FUNCTION_BLOCK FTS_NCGenerator
VAR_IN_OUT
	stAxis: ST_Axis;
END_VAR
VAR_INPUT
	///滤波窗口大小
	nWindowSize: UINT;
	fCycleTime: LREAL;
END_VAR
VAR
	///_bCalStart             :BOOL:=FALSE;
	_bEnable: BOOL;
	///_bAutoPlan             :BOOL:=FALSE;
	_bCalculateDone: BOOL;
	_bSynMode: BOOL := FALSE;
	_bFisrtUpdate: BOOL := FALSE;
	_bEndOfProfile: BOOL := FALSE;
	_bEstopping: BOOL := FALSE;
	///03.31     
	_bIsGroupMember: BOOL := FALSE;
	_bAddNodeOk: BOOL := FALSE;
	_bDeleteNodeOk: BOOL := FALSE;
	_bInsertOk: BOOL := FALSE;
	_bPreEstop  :BOOL:=FALSE;
	_bPreDyEstop  :BOOL:=FALSE;
	_nIndex: INT;
	_nNodeIndex: UINT;
	_nLastIndex: INT;
	_nPointIndex: UINT;
	_nForwardIndex: INT;
	_nPreIndex: INT;
	_nState: INT;
	_nPathSegment: INT;
	_nSysType: UINT;
	_nCamBufferNum: UINT := 0;
	_nCuRoadID: UINT;
	_nLastRoadID: UINT;
	_nMoverCounter: UINT;
	_nLastMoverCounter: UINT;
	_fRealDis: LREAL;
	_fPos: LREAL;
	_fSynPos: LREAL;
	_fSynVelo: LREAL;
	_lastVelo: LREAL;
	_fVeloStart: LREAL;
	_fVeloEnd: LREAL;
	_fTargetVelo: LREAL;
	_fStartPos: LREAL;
	_fEndPos: LREAL;
	_fVeloStart_2: LREAL;
	_fVeloEnd_2: LREAL;
	_fTargetVelo_2: LREAL;
	_fDistance_2: LREAL;
	_fAcc: LREAL;
	_fDec: LREAL;
	_fJerk: LREAL;
	_fAcc_2: LREAL;
	_fDec_2: LREAL;
	_fDistance: LREAL;
	///_fDistance_2             :LREAL;
	_fSetVelo: LREAL;
	///夹具长度*0.5
	_fGap: LREAL;
	_fGapSet: LREAL;
	_fTime: LREAL;
	_fDisSet: LREAL;
	_fForwardTime: LREAL;
	_fDealtDis: LREAL;
	_fDealt_S: LREAL;
	_fPre_S: LREAL;
	_fPreDealt_S: LREAL;
	_fDealt_S1: LREAL;
	_fPreCuVel: LREAL;
	_fCuVel: LREAL;
	_fPreTaVel: LREAL;
	_fPreAcc: LREAL;
	_fNewAcc: LREAL;
	_fDecTime: LREAL;
	_fDecTime_1: LREAL;
	_fPreCurTime: LREAL;
	_fPreSeg1TotalTime: LREAL;
	_fDisDiff: LREAL;
	_fDealDecTime: LREAL;
	_fMinDis: LREAL;
	_fNewAccDis: LREAL;
	_fReminDis: LREAL;
	_fAccMisDis: LREAL;
	_fAccMisDis_1: LREAL;
	_fNewVelo: LREAL;
	_fStartLinearPos: LREAL;
	_fLinearDealt: LREAL;
	_fMasterPos: LREAL;
	_fMasterStartPos: LREAL;
	_fMasterEndPos: LREAL;
	_fSlaveStartPos: LREAL;
	_fDePos: LREAL;
	_fDeCuVelo: LREAL;
	_fVeloRatio: LREAL;
	_fPos_X: LREAL;
	_fDealt_X: LREAL;
	_fLastPos: LREAL;
	_fMasterGap: LREAL;
	_fRoad1_Lenth: LREAL;
	_fRoad2_Lenth: LREAL;
	_fCuRoadLenth: LREAL;
	_fPosTemp: LREAL;
	_fLastPosDeat: LREAL;
	_fLastPosNC: LREAL;
	_fPosIn: LREAL;
	_fStopPos: LREAL;
	_fEStopPos: LREAL;
	_fPreStopPos: LREAL;
	_fUpNewPos: LREAL;
	_fUpNewPosTemp: LREAL;
	/// 成组组内gap 03.31
	_fGroupInGap: LREAL;
	///06.30
	_fSetDealtGap: LREAL;
	_fPyRealdis  :LREAL; //02.28
	_fLastRoadPos :LREAL;
	_fBreakDis    :LREAL;   
	_fSetSafeDis  :LREAL;
	_fLastPtyPos  :LREAL;
	_fPtyVelo    :LREAL;
	
	_fPreDealtP  :LREAL;
	
	///_fEndPos               :LREAL;  //03.26
	_sMessage3: STRING;
	_sMessage: STRING(1024);
	_sMessage2: STRING(1024);
	
	_pPremover: POINTER TO ST_Axis;
	_pNextRoadPremover: POINTER TO ST_Axis;
	///_fStopTime             :LREAL;
	_ePlanningMode: E_PlanningMode;
	_stAxis_Point: ST_Point;
	_stLastAxis_Point: ST_Point;
	_stForwardAxis_Point: ST_Point;
	_stPreAxis_Point: ST_Point;
	_stAxisNo: ST_Axis;
	_eDirection: E_Direction;
	///04.08
	_eSetDirection: E_Direction;
	_stTimeInfo: ST_TimeRef;
	_stTimeInfo_2: ST_TimeRef;
	_stPathRef: ST_PathRef;
	_stNoPathRef: ST_PathRef;
	_stPolynom5Factor: ST_Polynom5Factor;
	_stSShapedParam: ST_SParam;
	_stCamParam: ST_CamParam;
	_aLinearPosition: ARRAY[1..100] OF LREAL;
	_aCamBuffer: ARRAY[0..9] OF ST_CamXYVA;
	_fbTrig: R_TRIG;
	_fbSlaveTrig: R_TRIG;
	_fbPathTrig: R_TRIG;
	_fbDecPathTrig: R_TRIG;
	_fbCamPointUpdateTrig: R_TRIG;
	_fbCamBufUpdateTrig: R_TRIG;
	_fbClearFtrig: F_TRIG;
	_fbDecNextPathTrig: R_TRIG;
	_fbAxis: FB_TrajectoryPlanning;
	_fbPreAxis: FB_TrajectoryPlanning;
	_fbTon: TON;
	_fbFilterV2: FB_FilterWindowV2;
	_fbStopTrig: R_TRIG;
	_fbStopTon: TON;
	_fbAxisGroupList: FTS_AxisGroupList;
	_fbTrigRoadUpdate: R_TRIG;
	_fbTrigRoadDeleUpdate: R_TRIG;
	_fbTonCuPos:ton ; //02.28
END_VAR
VAR CONSTANT
	//cDebug: BOOL := TRUE;
	cStateIdle: INT := 0;
	cStateReady: INT := 1;
	cStatePathGenerator: INT := 2;
	cDealtGap: REAL := 10000;
	//cNcCycle: REAL := 0.001;
	cPointBuffer: UINT := 10;
END_VAR


// control logic 
IF stAxis.stAxisStatus.bPositiveDirection THEN 
	_eDirection:=E_Direction.DIRECTION_POSITIVE;
	
ELSIF stAxis.stAxisStatus.bNegativeDirection  THEN
	_eDirection:=E_Direction.DIRECTION_NEGATIVE;
	
ELSE
	_eDirection:=E_Direction.DIRECTION_POSITIVE;
END_IF

//根据不同road 前置和后置配置  04/02
IF (stAxis.stPLCTONC.nRoadID_2<>0)AND (stAxis.stPLCTONC.nRoadID_1<>0)AND(stAxis.stNcTOPLC.nCuRoadID=stAxis.stPLCTONC.nRoadID_2)THEN   //04.02
	
		IF NOT stAxis.stPLCTONC.bRoadDirection  THEN
			IF (stAxis.stAxisStatus.pPremover=0)THEN 
				_pPremover:=ADR(_stAxisNo);
			ELSE
				_pPremover:=stAxis.stAxisStatus.pPremover;
			END_IF
		ELSE
			IF (stAxis.stAxisStatus.pAftermover=0)THEN 
				_pPremover:=ADR(_stAxisNo);
			ELSE
				_pPremover:=stAxis.stAxisStatus.pAftermover;
			END_IF
		END_IF	
ELSE
	IF (_eDirection=E_Direction.DIRECTION_POSITIVE)THEN 
		IF (stAxis.stAxisStatus.pPremover=0)THEN 
			_pPremover:=ADR(_stAxisNo);
		ELSE
			_pPremover:=stAxis.stAxisStatus.pPremover;
		END_IF
	ELSE
		IF (stAxis.stAxisStatus.pAftermover=0)THEN 
			_pPremover:=ADR(_stAxisNo);
		ELSE
			_pPremover:=stAxis.stAxisStatus.pAftermover;
		END_IF
	
	END_IF
END_IF

IF (stAxis.stAxisStatus.pNextRoadPremover=0)THEN
	_pNextRoadPremover :=ADR(_stAxisNo);
ELSE
	_pNextRoadPremover :=stAxis.stAxisStatus.pNextRoadPremover;
END_IF

// 是否成组判断，并根据条件计算组内gap距离  03.31
IF (_pPremover^.stNcTOPLC.nAxisId<>0) THEN 
	IF (_pPremover^.stAxisStatus.stGroupRef.eGroupType<>E_GroupType.GROUPTYPE_NONE)
           AND (stAxis.stAxisStatus.stGroupRef.eGroupType<>E_GroupType.GROUPTYPE_NONE)THEN 
		IF (_pPremover^.stAxisStatus.stGroupRef.nGroupId=stAxis.stAxisStatus.stGroupRef.nGroupId)THEN 
			//_fGroupInGap:=stAxis.stAxisStatus.stPathRef.fGroupInGap;
			_fGroupInGap:=stAxis.stPLCTONC.fGroupInGap;
			_bIsGroupMember:=TRUE;
		END_IF
	ELSE
		_bIsGroupMember:=FALSE;
	END_IF
ELSE
	IF (_pNextRoadPremover^.stNcTOPLC.nAxisId<>0) THEN 
		IF (_pNextRoadPremover^.stAxisStatus.stGroupRef.eGroupType<>E_GroupType.GROUPTYPE_NONE)
			   AND (stAxis.stAxisStatus.stGroupRef.eGroupType<>E_GroupType.GROUPTYPE_NONE)THEN 
			IF (_pNextRoadPremover^.stAxisStatus.stGroupRef.nGroupId=stAxis.stAxisStatus.stGroupRef.nGroupId)THEN 
				//_fGroupInGap:=stAxis.stAxisStatus.stPathRef.fGroupInGap;
				_fGroupInGap:=stAxis.stPLCTONC.fGroupInGap;
				_bIsGroupMember:=TRUE;
			END_IF
		ELSE
			_bIsGroupMember:=FALSE;
		END_IF
	ELSE 
	   _bIsGroupMember:=FALSE;
	END_IF
END_IF



// 前后动子实时位置计算
IF stAxis.stPLCTONC.bNcEnable THEN 
	//IF (_pPremover^.stNcTOPLC.nAxisId<>0)THEN   //04.11
	IF (_pPremover^.stNcTOPLC.nAxisId<>0)AND (stAxis.stNcTOPLC.nCuRoadID=_pPremover^.stNcTOPLC.nCuRoadID)THEN   //04.11
		IF (stAxis.stNcTOPLC.nCuRoadID<>stAxis.stPLCTONC.nRoadID_2)THEN   //04.02
		    IF (_eDirection=E_Direction.DIRECTION_POSITIVE)THEN
				 IF (_pPremover^.stNcTOPLC.fActPos<stAxis.stNcTOPLC.fActPos)AND(stAxis.stPLCTONC.nSysType=3)THEN
					 _fRealDis:=_pPremover^.stNcTOPLC.fActPos+stAxis.stNcTOPLC.fModuloFactor-stAxis.stNcTOPLC.fActPos;
				 ELSE
					 _fRealDis:=_pPremover^.stNcTOPLC.fActPos-stAxis.stNcTOPLC.fActPos;
					 //_fPyRealdis:=_pPremover^.stCodToNCParam.fActualPos-stAxis.stCodToNCParam.fActualPos;  
				 END_IF
			ELSE
				IF (_pPremover^.stNcTOPLC.fActPos>stAxis.stNcTOPLC.fActPos)AND(stAxis.stPLCTONC.nSysType=3)THEN  
					 _fRealDis:=stAxis.stNcTOPLC.fActPos+stAxis.stNcTOPLC.fModuloFactor-_pPremover^.stNcTOPLC.fActPos; 
				ELSE
					_fRealDis:=stAxis.stNcTOPLC.fActPos-_pPremover^.stNcTOPLC.fActPos;
					//_fPyRealdis:=stAxis.stCodToNCParam.fActualPos-_pPremover^.stCodToNCParam.fActualPos;    //02.28
				END_IF
			END_IF
			
		ELSE
			IF NOT stAxis.stPLCTONC.bRoadDirection  THEN
				 _fRealDis:=_pPremover^.stNcTOPLC.fActPos-stAxis.stNcTOPLC.fActPos;
				 //_fPyRealdis:=_pPremover^.stCodToNCParam.fActualPos-stAxis.stCodToNCParam.fActualPos;    //02.28
			ELSE
				_fRealDis:=stAxis.stNcTOPLC.fActPos-_pPremover^.stNcTOPLC.fActPos;
				//_fPyRealdis:=stAxis.stCodToNCParam.fActualPos-_pPremover^.stCodToNCParam.fActualPos;    //02.28
			END_IF
		END_IF
		
		_fGapSet:=_pPremover^.stAxisStatus.stPathRef.fGap+stAxis.stAxisStatus.stPathRef.fSetGap;
		
		IF _bIsGroupMember THEN   //03.31
			_fGapSet:=_fGroupInGap;
		END_IF
	ELSE    //02.20 增加下一路段实时距离计算
		//IF ( _pNextRoadPremover^.stNcTOPLC.nAxisId<>0)THEN   04/11
		IF ( _pNextRoadPremover^.stNcTOPLC.nAxisId<>0)AND (stAxis.stNcTOPLC.nCuRoadID<>stAxis.stPLCTONC.nRoadID_2)AND(stAxis.stPLCTONC.nRoadID_2<>0) THEN  // 04/11
			IF (_eDirection=E_Direction.DIRECTION_POSITIVE)THEN
				  IF NOT stAxis.stPLCTONC.bRoadDirection  THEN   //正向
				      _fRealDis:=FC_TransformPosition(fOffset:=stAxis.stPLCTONC.fRoad1_Length, fPosition:=_pNextRoadPremover^.stNcTOPLC.fActPos)-stAxis.stNcTOPLC.fActPos;
					 _fPyRealdis:=FC_TransformPosition(fOffset:=stAxis.stPLCTONC.fRoad1_Length, fPosition:=_pNextRoadPremover^.stCodToNCParam.fActualPos)-stAxis.stCodToNCParam.fActualPos;  //02.28
				  ELSE
				      _fRealDis:=FC_TransformPosition(fOffset:=stAxis.stPLCTONC.fRoad1_Length, fPosition:=stAxis.stPLCTONC.fRoad2_Length-_pNextRoadPremover^.stNcTOPLC.fActPos)-stAxis.stNcTOPLC.fActPos;
					  _fPyRealdis:=FC_TransformPosition(fOffset:=stAxis.stPLCTONC.fRoad1_Length, fPosition:=stAxis.stPLCTONC.fRoad2_Length-_pNextRoadPremover^.stCodToNCParam.fActualPos)-stAxis.stCodToNCParam.fActualPos;//02.28
				  END_IF
			ELSE
				IF NOT stAxis.stPLCTONC.bRoadDirection  THEN   //正向
				      _fRealDis:=_pNextRoadPremover^.stNcTOPLC.fActPos+stAxis.stNcTOPLC.fActPos;  //04.17
					  _fPyRealdis:=_pNextRoadPremover^.stCodToNCParam.fActualPos+stAxis.stCodToNCParam.fActualPos;  //02.28
				  ELSE
				      _fRealDis:=stAxis.stNcTOPLC.fActPos+stAxis.stPLCTONC.fRoad2_Length-_pNextRoadPremover^.stNcTOPLC.fActPos;  //04.17
					  _fPyRealdis:=stAxis.stCodToNCParam.fActualPos+stAxis.stPLCTONC.fRoad2_Length-_pNextRoadPremover^.stCodToNCParam.fActualPos;  //02.28
				  END_IF
				  
			END_IF
			_fGapSet:=_pNextRoadPremover^.stAxisStatus.stPathRef.fGap+stAxis.stAxisStatus.stPathRef.fSetGap;
			IF _bIsGroupMember THEN   //03.31
				_fGapSet:=_fGroupInGap;
			END_IF
		ELSE
			_fRealDis:=0;
		END_IF 
	END_IF
	// 实时位置计算  07.16
	IF (_pPremover^.stNcTOPLC.nAxisId<>0) THEN
       IF (stAxis.stCodToNCParam.nRoadID=_pPremover^.stCodToNCParam.nRoadID)THEN   //07.16
			_fPyRealdis:=ABS(stAxis.stCodToNCParam.fActualPos-_pPremover^.stCodToNCParam.fActualPos);
		ELSE
			IF (stAxis.stCodToNCParam.nRoadID=stAxis.stPLCTONC.nRoadID_1)THEN
				IF (_eDirection=E_Direction.DIRECTION_POSITIVE)THEN
					IF NOT stAxis.stPLCTONC.bRoadDirection  THEN
						_fPyRealdis:=stAxis.stPLCTONC.fRoad1_Length-stAxis.stCodToNCParam.fActualPos+_pPremover^.stCodToNCParam.fActualPos;
					ELSE
						_fPyRealdis:=stAxis.stPLCTONC.fRoad1_Length-stAxis.stCodToNCParam.fActualPos+stAxis.stPLCTONC.fRoad2_Length-_pPremover^.stCodToNCParam.fActualPos;
					END_IF
				ELSE
					IF NOT stAxis.stPLCTONC.bRoadDirection  THEN
						_fPyRealdis:=stAxis.stCodToNCParam.fActualPos+_pPremover^.stCodToNCParam.fActualPos;
					ELSE
						_fPyRealdis:=stAxis.stCodToNCParam.fActualPos+stAxis.stPLCTONC.fRoad2_Length-_pPremover^.stCodToNCParam.fActualPos;
					END_IF
				END_IF
     
        END_IF 
			
		END_IF  
	END_IF
	stAxis.stAxisStatus.nNcCycleCounter_WP:=stAxis.stAxisStatus.nNcCycleCounter_WP+1;
ELSE
	stAxis.stAxisStatus.nNcCycleCounter_WP:=0;
END_IF 

//  dealtGap预值设置  //06.30
(*IF stAxis.stPLCTONC.fDealtGap<>0THEN
   _fSetDealtGap:=stAxis.stPLCTONC.fDealtGap;
ELSE
	_fSetDealtGap:=cDealtGap ;
END_IF*)
_fSetDealtGap:=cDealtGap ;

CASE  _nState  OF 
	cStateIdle:
	
	      IF stAxis.stPLCTONC.bNcEnable THEN 
              _nState:=cStateReady;
          END_IF       

    cStateReady:     
	      A_NCStartCase();
		  IF _bEnable THEN 
			  _nState:=cStatePathGenerator;
			  A_Planning();
			  _bEnable:=FALSE;
			  _stPathRef.bCalculateDone:=FALSE;
		  END_IF
    cStatePathGenerator:
	     
	      _nState:=cStateReady;

END_CASE
 

IF stAxis.stPLCTONC.bNcEnable AND _bCalculateDone THEN 
	
    A_GetPosition();
ELSE
	_bEndOfProfile:=FALSE;
	stAxis.stNcTOPLC.fActVelo:=0;
	stAxis.stAxisStatus.nNcCycleCounter:=0;   //06.20
END_IF

IF stAxis.stAxisStatus.nNcCycleCounter=0 THEN   //10.28
	stAxis.stAxisStatus.bSynStopping:=FALSE;
	//stAxis.stAxisStatus.bEmStopping:=FALSE;     //03.03   通信时序问题？？？
	_bEstopping:=FALSE;
END_IF

// 位置滤波
A_PositionHandle();

//动子前置和后置更新
A_NodeUpdate();  //04.20

ACTION A_AccSegmengt:

_fPreTaVel:=_pPremover^.stAxisStatus.stPathRef.fTargetVelocity;
_fPreCuVel:=_pPremover^.stNcTOPLC.fActVelo;
_fPreAcc:=_pPremover^.stAxisStatus.stPathRef.aExecutablePath[0].fAccleration;   //有问题

_fCuVel:=stAxis.stNcTOPLC.fActVelo;

// 匀速段
(*IF (_fCuVel>=stAxis.stAxisStatus.stPathRef.fTargetVelocity)THEN   //速度>=目标速度
	_fDealt_S1:=0.5*(_fPreTaVel-_fPreCuVel)*(_fPreTaVel-_fPreCuVel)/_fAcc;				     			   
	_fNewAcc:=(_fCuVel-_fPreTaVel)*(_fCuVel-_fPreTaVel)*0.5/(_fDealt_S+_fDealt_S1);
					 
	_fDecTime:=	(_fCuVel-_fPreTaVel)/_fNewAcc;
	_fNewAccDis:=(_fCuVel*_fCuVel-_fPreTaVel*_fPreTaVel)*0.5/_fNewAcc;   //减速面积
	_fMinDis:=_fPreTaVel*_fPreTaVel*0.5/_fAcc+_fNewAccDis;  //减速面积+停止最小面积
	_fPos:=stAxis.stPLCTONC.stEndPosition.fPosition;
	IF(_fReminDis< _fMinDis)THEN
			_fVeloStart:=stAxis.stNcTOPLC.fActVelo;
			_fVeloEnd:=0.0;
			_fTargetVelo:=_pPremover^.stAxisStatus.stPathRef.fTargetVelocity;
			_fAcc:=stAxis.stPLCTONC.stEndPosition.fAccleration;
			_fDec:=stAxis.stPLCTONC.stEndPosition.fDeceleration;
			IF (_eDirection=E_Direction.DIRECTION_POSITIVE)THEN
				_fDistance:=_fPos-stAxis.stNcTOPLC.fActPos;
			ELSE
				_fDistance:=stAxis.stNcTOPLC.fActPos-_fPos;
			END_IF
			_fAcc:=stAxis.stPLCTONC.stEndPosition.fAccleration;
			_fDec:=stAxis.stPLCTONC.stEndPosition.fDeceleration;
			_nPathSegment:=1;
	ELSE
			_nPathSegment:=2;
			_fVeloStart:=stAxis.stNcTOPLC.fActVelo;
			_fVeloEnd:=_fPreTaVel;
			_fTargetVelo:=_fPreTaVel;
			_fDistance:=_fNewAccDis;
			_fAcc:=_fNewAcc;
			_fDec:=_fNewAcc;
			
			_fVeloStart_2:=_fPreTaVel;
			_fVeloEnd_2:=0.0;
			_fTargetVelo_2:=_fPreTaVel;
			IF (_eDirection=E_Direction.DIRECTION_POSITIVE)THEN
				_fDistance_2:=_fPos-stAxis.stNcTOPLC.fActPos-_fNewAccDis;
			ELSE
				_fDistance_2:=stAxis.stNcTOPLC.fActPos-_fPos-_fNewAccDis;
			END_IF
			_fAcc_2:=stAxis.stPLCTONC.stEndPosition.fAccleration;
			_fDec_2:=stAxis.stPLCTONC.stEndPosition.fDeceleration;
			
	END_IF
	
	_bSynMode:=TRUE;
	_bEnable:=TRUE;
ELSIF (_fCuVel>=_fPreTaVel) THEN   //速度>前动子目标速度
	//_fAccMisDis:=0.5*(stAxis.stAxisStatus.stPathRef.fTargetVelocity-_fPreTaVel)*(stAxis.stAxisStatus.stPathRef.fTargetVelocity-_fPreTaVel)/_fAcc;
	_fAccMisDis:=(stAxis.stAxisStatus.stPathRef.fTargetVelocity-_fPreTaVel)*(stAxis.stAxisStatus.stPathRef.fTargetVelocity-_fPreTaVel)/_fAcc;
	_fDealt_S1:=0.5*(_fPreTaVel-_fPreCuVel)*(_fPreTaVel-_fPreCuVel)/_fAcc;
    IF(_fAccMisDis>=(_fDealt_S+_fDealt_S1)) THEN
		_fNewVelo:=_fPreTaVel+SQRT((_fDealt_S+_fDealt_S1)*_fAcc);
		_fNewAccDis:=(_fNewVelo*_fNewVelo-_fPreTaVel*_fPreTaVel)/_fAcc;  //减速追击面积
		//_fMinDis:=_fPreTaVel*_fPreTaVel*0.5/_fAcc+_fAccMisDis+_fNewAccDis;
		
		_fMinDis:=_fPreTaVel*_fPreTaVel*0.5/_fAcc+_fNewAccDis;
		IF(_fReminDis>=_fMinDis)THEN
			_nPathSegment:=2;
			_fVeloStart:=stAxis.stNcTOPLC.fActVelo;
			_fVeloEnd:=_fPreTaVel;
			_fTargetVelo:=_fNewVelo;
			_fDistance:=_fNewAccDis;
			_fAcc:=stAxis.stPLCTONC.stEndPosition.fAccleration;
			_fDec:=stAxis.stPLCTONC.stEndPosition.fDeceleration;
			
			_fVeloStart_2:=_fPreTaVel;
			_fVeloEnd_2:=0.0;
			_fTargetVelo_2:=_fPreTaVel;
			IF (_eDirection=E_Direction.DIRECTION_POSITIVE)THEN
				_fDistance_2:=_fPos-stAxis.stNcTOPLC.fActPos-_fNewAccDis;
			ELSE
				_fDistance_2:=stAxis.stNcTOPLC.fActPos-_fPos-_fNewAccDis;
			END_IF
			_fAcc_2:=stAxis.stPLCTONC.stEndPosition.fAccleration;
			_fDec_2:=stAxis.stPLCTONC.stEndPosition.fDeceleration;
			
	    END_IF
	
	END_IF

ELSE     //  其他情况不处理
    RETURN;
END_IF*)
IF (_fCuVel>_fPreTaVel)THEN   //速度>前动子目标速度
	    _fDealt_S1:=0.5*(_fPreTaVel-_fPreCuVel)*(_fPreTaVel-_fPreCuVel)/_fAcc;	
		
        IF (_fDealt_S>_fDealt_S1)THEN	   
	         _fNewAcc:=(_fCuVel-_fPreTaVel)*(_fCuVel-_fPreTaVel)*0.5/(_fDealt_S-_fDealt_S1);
			 IF (_fNewAcc>stAxis.stAxisParam.stDynamicDefault.fMaxDeceleration)THEN 
			    _fNewAcc:=stAxis.stAxisParam.stDynamicDefault.fMaxDeceleration;
		     END_IF
		ELSE
			_fNewAcc:=stAxis.stAxisParam.stDynamicDefault.fMaxDeceleration;
		END_IF
		
	    _fDecTime:=	(_fCuVel-_fPreTaVel)/_fNewAcc;
	    _fNewAccDis:=(_fCuVel*_fCuVel-_fPreTaVel*_fPreTaVel)*0.5/_fNewAcc;   //减速面积
	    _fMinDis:=_fPreTaVel*_fPreTaVel*0.5/_fAcc+_fNewAccDis;  //减速面积+停止最小面积
	    _fPos:=stAxis.stPLCTONC.stEndPosition.fPosition;
	    IF(_fReminDis< _fMinDis)THEN
			_fVeloStart:=stAxis.stNcTOPLC.fActVelo;
			_fVeloEnd:=0.0;
			_fTargetVelo:=_pPremover^.stAxisStatus.stPathRef.fTargetVelocity;
			_fAcc:=stAxis.stPLCTONC.stEndPosition.fAccleration;
			_fDec:=stAxis.stPLCTONC.stEndPosition.fDeceleration;
			IF (_eDirection=E_Direction.DIRECTION_POSITIVE)THEN
				_fDistance:=_fPos-stAxis.stNcTOPLC.fActPos;
			ELSE
				_fDistance:=stAxis.stNcTOPLC.fActPos-_fPos;
			END_IF
			
			_nPathSegment:=1;
	    ELSE
			_nPathSegment:=2;
			_fVeloStart:=stAxis.stNcTOPLC.fActVelo;
			_fVeloEnd:=_fPreTaVel;
			_fTargetVelo:=_fPreTaVel;
			_fDistance:=_fNewAccDis;
			_fAcc:=_fNewAcc;
			_fDec:=_fNewAcc;
			_fPosIn:=_fDealt_S;       
			_fVeloStart_2:=_fPreTaVel;
			_fVeloEnd_2:=0.0;
			_fTargetVelo_2:=_fPreTaVel;
			IF (_eDirection=E_Direction.DIRECTION_POSITIVE)THEN
				_fDistance_2:=_fPos-stAxis.stNcTOPLC.fActPos-_fNewAccDis;
			ELSE
				_fDistance_2:=stAxis.stNcTOPLC.fActPos-_fPos-_fNewAccDis;
			END_IF
			_fAcc_2:=stAxis.stPLCTONC.stEndPosition.fAccleration;
			_fDec_2:=stAxis.stPLCTONC.stEndPosition.fDeceleration;	
	   END_IF
	
ELSE     //按当前速度重新规划
	        (*_fVeloStart:=stAxis.stNcTOPLC.fActVelo;
			_fVeloEnd:=0.0;
			_fTargetVelo:=stAxis.stNcTOPLC.fActVelo;
			_fAcc:=stAxis.stPLCTONC.stEndPosition.fAccleration;
			_fDec:=stAxis.stPLCTONC.stEndPosition.fDeceleration;
			IF (_eDirection=E_Direction.DIRECTION_POSITIVE)THEN
				_fDistance:=_fPos-stAxis.stNcTOPLC.fActPos;
			ELSE
				_fDistance:=stAxis.stNcTOPLC.fActPos-_fPos;
			END_IF
			
			_nPathSegment:=1;*)
		RETURN;
END_IF
_bSynMode:=TRUE;
_bEnable:=TRUE;
stAxis.stAxisStatus.bSynDecActive:=TRUE;
IF GVL_MC.cDebug  THEN
	_sMessage:=FC_StrContact(stAxis,'acc gap control');
	ADSLOGSTR(ADSLOG_MSGTYPE_HINT, _sMessage, '');
END_IF
END_ACTION

ACTION A_CatchUp:

//  追击
(***********
   1. 前后动子间距小于防碰撞距离return 
   2. 前后动子间距小于欲减速设置距离，触发减速
   3. 判断当前动子有几段路径，分路径讨论前动子处于路径第几段和处于第几段的加速段、减速段和匀速段

************)

IF (_pPremover^.stNcTOPLC.nAxisId<>0)AND (NOT _bSynMode) THEN 
	//预处理减速距离,前瞻距离
	_fDisSet:=0.5*stAxis.stAxisStatus.stPathRef.fTargetVelocity*stAxis.stAxisStatus.stPathRef.fTargetVelocity/_fAcc;        
	
	IF (_nPathSegment=1)THEN 
		IF(_fTime<stAxis.stAxisStatus.stPathRef.aExecutablePath[0].fTa)THEN     // 当前动子处于第一减速段
			IF (stAxis.stAxisStatus.stPathRef.aExecutablePath[0].fExpVelo<stAxis.stAxisStatus.stPathRef.aExecutablePath[0].fStartVelo)
				AND (stAxis.stAxisStatus.stPathRef.aExecutablePath[0].fTv<>0)  THEN
				 _fDisSet:=0.5*stAxis.stAxisStatus.stPathRef.aExecutablePath[0].fStartVelo*stAxis.stAxisStatus.stPathRef.aExecutablePath[0].fStartVelo/_fAcc;
			END_IF
			
		END_IF
	ELSIF(_nPathSegment=2)THEN 
		IF(_fTime<stAxis.stAxisStatus.stPathRef.aExecutablePath[0].fTa)THEN
		    _fDisSet:=0.5*stAxis.stAxisStatus.stPathRef.aExecutablePath[0].fStartVelo*stAxis.stAxisStatus.stPathRef.aExecutablePath[0].fStartVelo/_fAcc;
		ELSE
			_fDisSet:=0.5*stAxis.stAxisStatus.stPathRef.aExecutablePath[1].fExpVelo*stAxis.stAxisStatus.stPathRef.aExecutablePath[1].fExpVelo/_fAcc;
		END_IF
	ELSE
		;
	END_IF
	_fDealt_S:=_fRealDis-_fGapSet;    //两动子间实时位置偏差，包含gap

	//IF ((_fRealDis -_fGapSet)<=cDealtGap)AND(_pPremover^.stAxisStatus.stPathRef.fTargetVelocity <stAxis.stAxisStatus.stPathRef.fTargetVelocity) THEN    //10.18 
	IF ((_fRealDis -_fGapSet)<=_fSetDealtGap)AND(_pPremover^.stAxisStatus.stPathRef.fTargetVelocity <stAxis.stAxisStatus.stPathRef.fTargetVelocity) THEN    //10.18 
		_fPos:=stAxis.stPLCTONC.stEndPosition.fPosition;
		_fTargetVelo:=_pPremover^.stAxisStatus.stPathRef.fTargetVelocity;
		_fVeloStart:=stAxis.stNcTOPLC.fActVelo;
		_fVeloEnd:=0;
		_fAcc:=stAxis.stPLCTONC.stEndPosition.fAccleration;
		_fDec:=stAxis.stPLCTONC.stEndPosition.fDeceleration;
		IF (_eDirection=E_Direction.DIRECTION_POSITIVE)THEN
		     _fDistance:=_fPos-stAxis.stNcTOPLC.fActPos;
	    ELSE
			 _fDistance:=stAxis.stNcTOPLC.fActPos-_fPos;
	    END_IF
		_bEnable:=TRUE;
		_nPathSegment:=1;
		stAxis.stAxisStatus.bSynDecActive:=TRUE;
		RETURN;
	 END_IF   //11.22 增加
	
    _fReminDis:=ABS(stAxis.stPLCTONC.stEndPosition.fPosition-stAxis.stNcTOPLC.fActPos);   //剩余目标距离
	
	IF (_fDealt_S-_fDisSet<=0)THEN    //触发减速判断
		   //IF (_pPremover^.stAxisStatus.stPathRef.fTargetVelocity <stAxis.stAxisStatus.stPathRef.fTargetVelocity) THEN  //11.25注释
		   IF (stAxis.stNcTOPLC.fActVelo>_pPremover^.stNcTOPLC.fActVelo) THEN     //11.25修改
			   IF (_fReminDis>_fDisSet)THEN  //判断剩余距离是否满足撞击条件,小于不处理 ，考虑减速距离过长特殊场景
				    _fPreCurTime:=UDINT_TO_LREAL(_pPremover^.stAxisStatus.nNcCycleCounter)*fCycleTime;
			       IF (_pPremover^.stAxisStatus.stPathRef._nPathSegmentNum=1)THEN      //判断前动子只有一段路径
				  
					   IF (_fPreCurTime <_pPremover^.stAxisStatus.stPathRef.aExecutablePath[0].fTa)THEN      //加速段或减速第一段
						   IF (_pPremover^.stAxisStatus.stPathRef.aExecutablePath[0].fExpVelo>_pPremover^.stAxisStatus.stPathRef.aExecutablePath[0].fStartVelo)THEN
							   IF (stAxis.stAxisStatus.stPathRef.aExecutablePath[0].fTv<>0) THEN          //加速段
								   A_AccSegmengt();
							   END_IF 
						   ELSE    //减速段
							   IF(_pPremover^.stAxisStatus.stPathRef.aExecutablePath[0].fTv<>0)THEN 
								   A_DecSegment();
							   END_IF
						   END_IF
					   // 匀速段
					   ELSIF (_fPreCurTime <(_pPremover^.stAxisStatus.stPathRef.aExecutablePath[0].fTotalTime-_pPremover^.stAxisStatus.stPathRef.aExecutablePath[0].fTd))THEN
						   A_ConVeloSegment();
					   ELSE
						   //
						   RETURN ;  //不处理
					   END_IF
				   //第二段
				   ELSIF(_pPremover^.stAxisStatus.stPathRef._nPathSegmentNum=2)THEN
                       IF (_pPremover^.stAxisStatus.nSegIndex=0) THEN   //前动子在第一段
						    //IF (_fPreCurTime <_pPremover^.stAxisStatus.stPathRef.aExecutablePath[0].fTa)THEN      //加速段
							IF (_fPreCurTime <_pPremover^.stAxisStatus.stPathRef.aExecutablePath[0].fTotalTime)THEN      //减速段  11.29
								A_DecSegment_2();
							END_IF
					   ELSIF (_pPremover^.stAxisStatus.nSegIndex=1) THEN   //只处理匀速段
						   IF (_fPreCurTime <(_pPremover^.stAxisStatus.stPathRef.aExecutablePath[1].fTotalTime-_pPremover^.stAxisStatus.stPathRef.aExecutablePath[1].fTd))THEN
						       A_ConVeloSegment();
						   END_IF   
					   ELSE
						   ;
					   END_IF
					   // 第二段减速段不处理
				   
				   END_IF
			   ELSE    //判断剩余距离是否满足撞击条件,小于不处理 ，考虑减速距离过长特殊场景,
				   
				   RETURN ;
		       END_IF
		   END_IF
	END_IF
END_IF
END_ACTION

ACTION A_ContantVeloPosition:
stAxis.stAxisStatus.nNcCycleCounter:=stAxis.stAxisStatus.nNcCycleCounter+1;
IF stAxis.stAxisStatus.bPositiveDirection THEN
	stAxis.stNcTOPLC.fActPos:=stAxis.stNcTOPLC.fActVelo*fCycleTime+stAxis.stNcTOPLC.fActPos;
ELSE
	stAxis.stNcTOPLC.fActPos:=stAxis.stNcTOPLC.fActPos-stAxis.stNcTOPLC.fActVelo*fCycleTime;
END_IF
stAxis.stNcTOPLC.fSetVelo:=stAxis.stNcTOPLC.fActVelo;
stAxis.stNcTOPLC.fSetAcc:=0;
stAxis.stNcTOPLC.fSetJerk:=0;
END_ACTION

ACTION A_ConVeloSegment:

_fPreTaVel:=_pPremover^.stAxisStatus.stPathRef.fTargetVelocity;
_fPreCuVel:=_pPremover^.stNcTOPLC.fActVelo;
_fPreAcc:=_fAcc;
_fCuVel:=stAxis.stNcTOPLC.fActVelo;
//_fDealt_S1:=0.5*(_fPreTaVel-_fPreCuVel)*(_fPreTaVel-_fPreCuVel)/_fAcc;
				      
_fNewAcc:=(_fCuVel-_fPreTaVel)*(_fCuVel-_fPreTaVel)*0.5/_fDealt_S;
		   		 
_fDecTime:=	(_fCuVel-_fPreTaVel)/_fNewAcc;
_fNewAccDis:=(_fCuVel*_fCuVel-_fPreTaVel*_fPreTaVel)*0.5/_fNewAcc;
_fMinDis:=_fPreTaVel*_fPreTaVel*0.5/_fPreAcc+_fNewAccDis;

_fPos:=stAxis.stPLCTONC.stEndPosition.fPosition;
	
IF(_fReminDis< _fMinDis)THEN
		_fVeloStart:=stAxis.stNcTOPLC.fActVelo;
	    _fVeloEnd:=0.0;
	    _fTargetVelo:=_pPremover^.stAxisStatus.stPathRef.fTargetVelocity;
		IF (_eDirection=E_Direction.DIRECTION_POSITIVE)THEN
			_fDistance:=_fPos-stAxis.stNcTOPLC.fActPos;
		ELSE
			_fDistance:=stAxis.stNcTOPLC.fActPos-_fPos;
		END_IF
		_fAcc:=stAxis.stPLCTONC.stEndPosition.fAccleration;
	    _fDec:=stAxis.stPLCTONC.stEndPosition.fDeceleration;
		_nPathSegment:=1;
ELSE
		_nPathSegment:=2;
		_fVeloStart:=stAxis.stNcTOPLC.fActVelo;
	    _fVeloEnd:=_fPreTaVel;
	    _fTargetVelo:=_fPreTaVel;
		_fDistance:=_fNewAccDis;
		_fAcc:=_fNewAcc;
	    _fDec:=_fNewAcc;
		_fPosIn:=_fDealt_S;       //11.29
	    _fVeloStart_2:=_fPreTaVel;
	    _fVeloEnd_2:=0.0;
	    _fTargetVelo_2:=_fPreTaVel;
		IF (_eDirection=E_Direction.DIRECTION_POSITIVE)THEN
			_fDistance_2:=_fPos-stAxis.stNcTOPLC.fActPos-_fNewAccDis;
		ELSE
			_fDistance_2:=stAxis.stNcTOPLC.fActPos-_fPos-_fNewAccDis;
		END_IF
		_fAcc_2:=stAxis.stPLCTONC.stEndPosition.fAccleration;
	    _fDec_2:=stAxis.stPLCTONC.stEndPosition.fDeceleration;
END_IF

_bSynMode:=TRUE;
_bEnable:=TRUE;
stAxis.stAxisStatus.bSynDecActive:=TRUE;
                
IF GVL_MC.cDebug  THEN
    _sMessage:=FC_StrContact(stAxis,'con gap control');
	 ADSLOGSTR(ADSLOG_MSGTYPE_HINT, _sMessage, '');
END_IF
END_ACTION

ACTION A_DecSegment:

_fPreTaVel:=_pPremover^.stAxisStatus.stPathRef.fTargetVelocity;
_fPreCuVel:=_pPremover^.stNcTOPLC.fActVelo;
_fPreAcc:=_fAcc;
_fCuVel:=stAxis.stNcTOPLC.fActVelo;

// 计算前动子的减速距离
_fPre_S:=(_fPreCuVel-_fPreTaVel)*(_fPreCuVel-_fPreTaVel)*0.5/_pPremover^.stAxisStatus.stPathRef.aExecutablePath[0].fDeceleration;
		      	   
//_fNewAcc:=(_fCuVel-_fPreTaVel)*(_fCuVel-_fPreTaVel)*0.5/_fDealt_S;  //06.18 
_fNewAcc:=(_fCuVel-_fPreTaVel)*(_fCuVel-_fPreTaVel)*0.5/(_fDealt_S+_fPre_S);  //06.18

//_fNewAcc:=(_fCuVel-_fPreTaVel)*(_fCuVel-_fPreTaVel)*0.5/_fDealt_S;
_fDecTime:=	(_fCuVel-_fPreTaVel)/_fNewAcc;
_fNewAccDis:=(_fCuVel*_fCuVel-_fPreTaVel*_fPreTaVel)*0.5/_fNewAcc;
_fMinDis:=_fPreTaVel*_fPreTaVel*0.5/_fPreAcc+_fNewAccDis;

_fPos:=stAxis.stPLCTONC.stEndPosition.fPosition;

IF(_fReminDis< _fMinDis)THEN
		_fVeloStart:=stAxis.stNcTOPLC.fActVelo;
	    _fVeloEnd:=0.0;
	    _fTargetVelo:=_pPremover^.stAxisStatus.stPathRef.fTargetVelocity;
		IF (_eDirection=E_Direction.DIRECTION_POSITIVE)THEN
			_fDistance:=_fPos-stAxis.stNcTOPLC.fActPos;
		ELSE
			_fDistance:=stAxis.stNcTOPLC.fActPos-_fPos;
		END_IF
		_fAcc:=stAxis.stPLCTONC.stEndPosition.fAccleration;
	    _fDec:=stAxis.stPLCTONC.stEndPosition.fDeceleration;
		_nPathSegment:=1;
ELSE
		_nPathSegment:=2;
		_fVeloStart:=stAxis.stNcTOPLC.fActVelo;
	    _fVeloEnd:=_fPreTaVel;
	    _fTargetVelo:=_fPreTaVel;
		_fDistance:=_fNewAccDis;
		_fAcc:=_fNewAcc;
	    _fDec:=_fNewAcc;
		
	    _fVeloStart_2:=_fPreTaVel;
	    _fVeloEnd_2:=0.0;
	    _fTargetVelo_2:=_fPreTaVel;
		_fPosIn:=_fDealt_S;       // 25.01.17
		IF (_eDirection=E_Direction.DIRECTION_POSITIVE)THEN
			_fDistance_2:=_fPos-stAxis.stNcTOPLC.fActPos-_fNewAccDis;
		ELSE
			_fDistance_2:=stAxis.stNcTOPLC.fActPos-_fPos-_fNewAccDis;
		END_IF
		_fAcc_2:=stAxis.stPLCTONC.stEndPosition.fAccleration;
	    _fDec_2:=stAxis.stPLCTONC.stEndPosition.fDeceleration;
END_IF
_bSynMode:=TRUE;
_bEnable:=TRUE;
stAxis.stAxisStatus.bSynDecActive:=TRUE;

IF GVL_MC.cDebug  THEN
		_sMessage:=FC_StrContact(stAxis,'dec gap control');
	     ADSLOGSTR(ADSLOG_MSGTYPE_HINT, _sMessage, '');
END_IF
END_ACTION

ACTION A_DecSegment_2:

_fPreTaVel:=_pPremover^.stAxisStatus.stPathRef.fTargetVelocity;
_fPreCuVel:=_pPremover^.stNcTOPLC.fActVelo;
_fPreAcc:=_fAcc;
_fCuVel:=stAxis.stNcTOPLC.fActVelo;
 _fPreSeg1TotalTime :=_pPremover^.stAxisStatus.stPathRef.aExecutablePath[0].fTotalTime;   //05.26
//_fPreDealt_S:=0.5*(_pPremover^.stAxisStatus.stPathRef.aExecutablePath[0].fTa-_fPreCurTime)*_fPreCuVel;
//_fPreDealt_S:=_pPremover^.stAxisStatus.stPathRef.fDealtInPos- 0.5*(_fPreTaVel+_fPreCuVel)*_fPreCurTime; //05.26  
_fPreDealt_S:=0.5*(_fPreCuVel-_fPreTaVel)*( _fPreSeg1TotalTime-_fPreCurTime); //05.26 
			      	   
_fNewAcc:=(_fCuVel-_fPreTaVel)*(_fCuVel-_fPreTaVel)*0.5/(_fDealt_S+_fPreDealt_S);
		   		 
_fDecTime:=	(_fCuVel-_fPreTaVel)/_fNewAcc;
_fNewAccDis:=(_fCuVel*_fCuVel-_fPreTaVel*_fPreTaVel)*0.5/_fNewAcc;

_fMinDis:=_fPreTaVel*_fPreTaVel*0.5/_fPreAcc+_fNewAccDis;

_fPos:=stAxis.stPLCTONC.stEndPosition.fPosition;

IF( _fReminDis< _fMinDis)THEN
		_fVeloStart:=stAxis.stNcTOPLC.fActVelo;
	    _fVeloEnd:=0.0;
	    _fTargetVelo:=_pPremover^.stAxisStatus.stPathRef.fTargetVelocity;
		IF (_eDirection=E_Direction.DIRECTION_POSITIVE)THEN
			_fDistance:=_fPos-stAxis.stNcTOPLC.fActPos;
		ELSE
			_fDistance:=stAxis.stNcTOPLC.fActPos-_fPos;
		END_IF
		_nPathSegment:=1;
		_fAcc:=stAxis.stPLCTONC.stEndPosition.fAccleration;
	    _fDec:=stAxis.stPLCTONC.stEndPosition.fDeceleration;
ELSE
		_nPathSegment:=2;
		_fVeloStart:=stAxis.stNcTOPLC.fActVelo;
	    _fVeloEnd:=_fPreTaVel;
	    _fTargetVelo:=_fPreTaVel;
		_fDistance:=_fNewAccDis;
		_fAcc:=_fNewAcc;
	    _fDec:=_fNewAcc;
		_fPosIn:=_fDealt_S+_fPreDealt_S;       //11.29
	    _fVeloStart_2:=_fPreTaVel;
	    _fVeloEnd_2:=0.0;
	    _fTargetVelo_2:=_fPreTaVel;
		IF (_eDirection=E_Direction.DIRECTION_POSITIVE)THEN
			_fDistance_2:=_fPos-stAxis.stNcTOPLC.fActPos-_fNewAccDis;
		ELSE
			_fDistance_2:=stAxis.stNcTOPLC.fActPos-_fPos-_fNewAccDis;
		END_IF
		_fAcc_2:=stAxis.stPLCTONC.stEndPosition.fAccleration;
	    _fDec_2:=stAxis.stPLCTONC.stEndPosition.fDeceleration;
		
END_IF
_bSynMode:=TRUE;
_bEnable:=TRUE;
stAxis.stAxisStatus.bSynDecActive:=TRUE;

IF GVL_MC.cDebug  THEN
		_sMessage:=FC_StrContact(stAxis,'dec2 gap control');
	     ADSLOGSTR(ADSLOG_MSGTYPE_HINT, _sMessage, '');
END_IF
END_ACTION

ACTION A_EStop:

//计算最小制动距离
_fPtyVelo:= ABS(_fLastPtyPos-stAxis.stCodToNCParam.fActualPos)/fCycleTime;  //实际速度
_fBreakDis:=0.5*stAxis.stNcTOPLC.fActVelo/(GVL_MC.nMaxDecRatio*stAxis.stPLCTONC.stEndPosition.fDeceleration);
//_fSetSafeDis:=UDINT_TO_LREAL(GVL_MC.nMecReserveDis+GVL_MC.nFollowError);
_fSetSafeDis:=UDINT_TO_LREAL(GVL_MC.nMecReserveDis);

// 07.14 增加前动子跟随误差计算  分两种情况判断 前动子停止 和运行两种状态
IF (_pPremover^.stNcTOPLC.nAxisId<>0)AND(stAxis.stAxisStatus.nNcCycleCounter<>0)THEN 
	_fPreDealtP :=ABS(_pPremover^.stNcTOPLC.fActPos-_pPremover^.stCodToNCParam.fActualPos);
	IF _fPreDealtP>GVL_MC.nFollowError AND _pPremover^.stAxisStatus.nNcCycleCounter<>0 THEN 
		_bPreDyEstop:=TRUE;
	ELSE
		_bPreDyEstop:=FALSE;
	END_IF 
	IF _pPremover^.stAxisStatus.nNcCycleCounter=0 THEN
		_bPreEstop:=TRUE;
	ELSE
		_bPreEstop:=FALSE;
	END_IF
    
ELSIF(_pNextRoadPremover^.stNcTOPLC.nAxisId<>0)AND(stAxis.stAxisStatus.nNcCycleCounter<>0) THEN
	IF (_pNextRoadPremover^.stNcTOPLC.nCuRoadID=_pNextRoadPremover^.stCodToNCParam.nRoadID)THEN
	    _fPreDealtP :=ABS(_pNextRoadPremover^.stNcTOPLC.fActPos-_pNextRoadPremover^.stCodToNCParam.fActualPos);
	ELSE
		IF (_eDirection=E_Direction.DIRECTION_POSITIVE)THEN
			IF NOT stAxis.stPLCTONC.bRoadDirection  THEN   //正向
				_fPreDealtP:=ABS(stAxis.stPLCTONC.fRoad1_Length+_pNextRoadPremover^.stNcTOPLC.fActPos-_pNextRoadPremover^.stCodToNCParam.fActualPos);
			ELSE
				_fPreDealtP:=ABS(stAxis.stPLCTONC.fRoad1_Length+stAxis.stPLCTONC.fRoad2_Length-_pNextRoadPremover^.stNcTOPLC.fActPos-_pNextRoadPremover^.stCodToNCParam.fActualPos);
			END_IF
		ELSE
			IF NOT stAxis.stPLCTONC.bRoadDirection  THEN   //正向
				_fPreDealtP:=ABS(_pNextRoadPremover^.stNcTOPLC.fActPos+_pNextRoadPremover^.stCodToNCParam.fActualPos);
			ELSE
				_fPreDealtP:=ABS(stAxis.stPLCTONC.fRoad2_Length-_pNextRoadPremover^.stNcTOPLC.fActPos+_pNextRoadPremover^.stCodToNCParam.fActualPos);
			END_IF
		
		END_IF
	END_IF
	
	IF _fPreDealtP>GVL_MC.nFollowError AND _pNextRoadPremover^.stAxisStatus.nNcCycleCounter<>0 THEN 
		_bPreDyEstop:=TRUE;
	ELSE
		_bPreDyEstop:=FALSE;
	END_IF 
	IF _pNextRoadPremover^.stAxisStatus.nNcCycleCounter=0 THEN
		_bPreEstop:=TRUE;
	ELSE
		_bPreEstop:=FALSE;
	END_IF
ELSE
	_fPreDealtP :=0;
	_bPreDyEstop:=FALSE;
	_bPreEstop:=FALSE;
END_IF

_fbTonCuPos(IN:=(_fPyRealdis<(_fGapSet-_fSetSafeDis)AND GVL_MC.bEmStop AND(_bPreEstop OR _bPreDyEstop)), PT:=T#10MS, Q=> , ET=> );  //06.22


IF _fRealDis<=0 OR _fPyRealdis<0  THEN  //02.28
	return;
END_IF

// 规划位置急停
IF (_pPremover^.stNcTOPLC.nAxisId<>0)AND (stAxis.stAxisStatus.nNcCycleCounter<>0)AND (_pPremover^.stNcTOPLC.nCuRoadID=stAxis.stNcTOPLC.nCuRoadID)  THEN  //04.08
	
	_fEStopPos:= 0.5*stAxis.stNcTOPLC.fActVelo*stAxis.stNcTOPLC.fActVelo/(GVL_MC.nMaxDecRatio*stAxis.stPLCTONC.stEndPosition.fDeceleration);  //07.13
	IF (_pPremover^.stAxisStatus.nNcCycleCounter=0) THEN
		IF _fRealDis <(_fGapSet-cDealtGap)  AND NOT _bEstopping  THEN   //11.06
                   IF (_eDirection=E_Direction.DIRECTION_POSITIVE)THEN    			  
	                    _fPos:=_fEStopPos+stAxis.stNcTOPLC.fActPos;
						//IF (stAxis.stPLCTONC.eCommand<>E_Command.COMMAND_ABSOLUTEFORK) THEN
						IF (stAxis.stPLCTONC.nRoadID_1=0)THEN 
							IF (_fPos>stAxis.stPLCTONC.fTargetPos)THEN     //03.20
								RETURN;
							END_IF
						ELSE  //驳指令
							IF (stAxis.stNcTOPLC.nCuRoadID=stAxis.stPLCTONC.nRoadID_1) THEN 
							   stAxis.stPLCTONC.stStartPosition.nRoadID:=stAxis.stPLCTONC.nRoadID_1;
							   stAxis.stPLCTONC.stEndPosition.nRoadID:=stAxis.stPLCTONC.nRoadID_1;
							   IF (_fPos>stAxis.stPLCTONC.fTargetPos)THEN     //03.20
								   RETURN;
							   END_IF
						    ELSE
							   stAxis.stPLCTONC.stStartPosition.nRoadID:=stAxis.stPLCTONC.nRoadID_2;
							   stAxis.stPLCTONC.stEndPosition.nRoadID:=stAxis.stPLCTONC.nRoadID_2;
							   IF NOT stAxis.stPLCTONC.bRoadDirection  THEN   //正向 
								    IF (_fPos>stAxis.stPLCTONC.fTargetPos)THEN     //03.20
								        RETURN;
							        END_IF
							   ELSE
								   IF (_fPos<stAxis.stPLCTONC.fTargetPos)THEN     //03.20
								        RETURN;
							       END_IF
							   END_IF
						    END_IF
							
						END_IF
				   ELSE
					    _fPos:=stAxis.stNcTOPLC.fActPos-_fEStopPos;
						
						//IF (stAxis.stPLCTONC.eCommand<>E_Command.COMMAND_ABSOLUTEFORK) THEN
						IF (stAxis.stPLCTONC.nRoadID_1=0)THEN 
							IF (_fPos<stAxis.stPLCTONC.fTargetPos)THEN     //03.20
								RETURN;
							END_IF
						ELSE  //非接驳指令
							IF (stAxis.stNcTOPLC.nCuRoadID=stAxis.stPLCTONC.nRoadID_1) THEN 
							   stAxis.stPLCTONC.stStartPosition.nRoadID:=stAxis.stPLCTONC.nRoadID_1;
							   stAxis.stPLCTONC.stEndPosition.nRoadID:=stAxis.stPLCTONC.nRoadID_1;
							   IF (_fPos<stAxis.stPLCTONC.fTargetPos)THEN     //03.20
								   RETURN;
							   END_IF
						    ELSE
							   stAxis.stPLCTONC.stStartPosition.nRoadID:=stAxis.stPLCTONC.nRoadID_2;
							   stAxis.stPLCTONC.stEndPosition.nRoadID:=stAxis.stPLCTONC.nRoadID_2;
							   IF NOT stAxis.stPLCTONC.bRoadDirection  THEN   //正向 
								    IF (_fPos>stAxis.stPLCTONC.fTargetPos)THEN     //03.20
								        RETURN;
							        END_IF
							   ELSE
								   IF (_fPos<stAxis.stPLCTONC.fTargetPos)THEN     //03.20
								        RETURN;
							       END_IF
							   END_IF
						    END_IF
							
						END_IF
				   END_IF
				   
				   _fTargetVelo:=stAxis.stNcTOPLC.fActVelo;
				   _fVeloStart:=stAxis.stNcTOPLC.fActVelo;
				   _fVeloEnd:=0;
				  // _fAcc:=stAxis.stAxisParam.stDynamicDefault.fMaxDeceleration;  //07.13
				  // _fDec:=stAxis.stAxisParam.stDynamicDefault.fMaxDeceleration;  //07.13
				   _fAcc:=GVL_MC.nMaxDecRatio*stAxis.stPLCTONC.stEndPosition.fAccleration;  //07.13
				   _fDec:=GVL_MC.nMaxDecRatio*stAxis.stPLCTONC.stEndPosition.fDeceleration; //07.13
				   
				   _fDistance:=_fEStopPos;
				   _bEnable:=TRUE;
				   _nPathSegment:=1;
				  // stAxis.stAxisStatus.bSynDecActive:=TRUE;
				   stAxis.stAxisStatus.bSynStopping:=TRUE;
		           _bEstopping:=TRUE;  
				 IF GVL_MC.cDebug  THEN
					_sMessage:=FC_StrContact(stAxis,'pPremover Estop path');
					 ADSLOGSTR(ADSLOG_MSGTYPE_HINT, _sMessage, '');
				END_IF
		END_IF
		
	END_IF
	
ELSE
	IF (_pNextRoadPremover^.stNcTOPLC.nAxisId<>0)AND (stAxis.stAxisStatus.nNcCycleCounter<>0) THEN 
		_fEStopPos:= 0.5*stAxis.stNcTOPLC.fActVelo*stAxis.stNcTOPLC.fActVelo/(GVL_MC.nMaxDecRatio*stAxis.stPLCTONC.stEndPosition.fDeceleration);  //07.13
		IF (_pNextRoadPremover^.stAxisStatus.nNcCycleCounter=0) THEN
			IF _fRealDis <(_fGapSet-cDealtGap) AND  NOT _bEstopping THEN  //11.06
				IF (_eDirection=E_Direction.DIRECTION_POSITIVE)THEN
					_fPos:=_fEStopPos+stAxis.stNcTOPLC.fActPos;
					IF (stAxis.stNcTOPLC.fActPos+_fEStopPos)>_fRoad1_Lenth THEN
						stAxis.stPLCTONC.stStartPosition.nRoadID:=stAxis.stPLCTONC.nRoadID_1;
						stAxis.stPLCTONC.stEndPosition.nRoadID:=stAxis.stPLCTONC.nRoadID_2;
                         IF NOT stAxis.stPLCTONC.bRoadDirection  THEN   //正向 
								 IF (_fPos>stAxis.stPLCTONC.fTargetPos)THEN     //03.20
								      RETURN;
							     END_IF
					     ELSE
								 IF (_fPos<stAxis.stPLCTONC.fTargetPos)THEN     //03.20
								        RETURN;
							     END_IF
					     END_IF
						
					ELSE
						stAxis.stPLCTONC.stStartPosition.nRoadID:=stAxis.stPLCTONC.nRoadID_1;
						stAxis.stPLCTONC.stEndPosition.nRoadID:=stAxis.stPLCTONC.nRoadID_1; 
					END_IF
			    ELSE
			        _fPos:=stAxis.stNcTOPLC.fActPos-_fEStopPos;
					IF (stAxis.stNcTOPLC.fActPos-_fStopPos)<0 THEN
						stAxis.stPLCTONC.stStartPosition.nRoadID:=stAxis.stPLCTONC.nRoadID_1;
						stAxis.stPLCTONC.stEndPosition.nRoadID:=stAxis.stPLCTONC.nRoadID_2; 
						IF NOT stAxis.stPLCTONC.bRoadDirection  THEN   //正向 
							IF (_fPos>stAxis.stPLCTONC.fTargetPos)THEN     //03.20
									  RETURN;
							 END_IF
						ELSE
							IF (_fPos<stAxis.stPLCTONC.fTargetPos)THEN     //03.20
									  RETURN;
							END_IF
					    END_IF
						
					ELSE
						stAxis.stPLCTONC.stStartPosition.nRoadID:=stAxis.stPLCTONC.nRoadID_1;
						stAxis.stPLCTONC.stEndPosition.nRoadID:=stAxis.stPLCTONC.nRoadID_1; 
					END_IF
					
			   END_IF 
			    _fDistance:=_fEStopPos;
                	
				_fAcc:=GVL_MC.nMaxDecRatio*stAxis.stPLCTONC.stEndPosition.fAccleration;  //07.13
				_fDec:=GVL_MC.nMaxDecRatio*stAxis.stPLCTONC.stEndPosition.fDeceleration; //07.13	
				_fTargetVelo:=stAxis.stNcTOPLC.fActVelo;
				_fVeloStart:=stAxis.stNcTOPLC.fActVelo;
				_fVeloEnd:=0;
				_bEnable:=TRUE;
				_nPathSegment:=1;
				stAxis.stAxisStatus.bSynStopping:=TRUE;
				_bEstopping:=TRUE;
				IF GVL_MC.cDebug  THEN
					_sMessage:=FC_StrContact(stAxis,'pNextRoadPremover Estop path');
					 ADSLOGSTR(ADSLOG_MSGTYPE_HINT, _sMessage, '');
				END_IF
			END_IF
	    END_IF			  	  
    END_IF
END_IF 

// 引入实际位置急停
IF (_pPremover^.stNcTOPLC.nAxisId<>0)AND (stAxis.stAxisStatus.nNcCycleCounter<>0)AND (_pPremover^.stNcTOPLC.nCuRoadID=stAxis.stNcTOPLC.nCuRoadID)  THEN  //04.08
	
	_fEStopPos:= 0.5*stAxis.stNcTOPLC.fActVelo*stAxis.stNcTOPLC.fActVelo/(GVL_MC.nMaxDecRatio*stAxis.stPLCTONC.stEndPosition.fDeceleration);  //07.13
	   IF _fbTonCuPos.Q  AND NOT _bEstopping  THEN   //02.28 增加实际距离检测
                   IF (_eDirection=E_Direction.DIRECTION_POSITIVE)THEN    			  
	                    _fPos:=_fEStopPos+stAxis.stNcTOPLC.fActPos;
						//IF (stAxis.stPLCTONC.eCommand<>E_Command.COMMAND_ABSOLUTEFORK) THEN
						IF (stAxis.stPLCTONC.nRoadID_1=0)THEN 
							IF (_fPos>stAxis.stPLCTONC.fTargetPos)THEN     //03.20
								RETURN;
							END_IF
						ELSE  //驳指令
							IF (stAxis.stNcTOPLC.nCuRoadID=stAxis.stPLCTONC.nRoadID_1) THEN 
							   stAxis.stPLCTONC.stStartPosition.nRoadID:=stAxis.stPLCTONC.nRoadID_1;
							   stAxis.stPLCTONC.stEndPosition.nRoadID:=stAxis.stPLCTONC.nRoadID_1;
							   IF (_fPos>stAxis.stPLCTONC.fTargetPos)THEN     //03.20
								   RETURN;
							   END_IF
						    ELSE
							   stAxis.stPLCTONC.stStartPosition.nRoadID:=stAxis.stPLCTONC.nRoadID_2;
							   stAxis.stPLCTONC.stEndPosition.nRoadID:=stAxis.stPLCTONC.nRoadID_2;
							   IF NOT stAxis.stPLCTONC.bRoadDirection  THEN   //正向 
								    IF (_fPos>stAxis.stPLCTONC.fTargetPos)THEN     //03.20
								        RETURN;
							        END_IF
							   ELSE
								   IF (_fPos<stAxis.stPLCTONC.fTargetPos)THEN     //03.20
								        RETURN;
							       END_IF
							   END_IF
						    END_IF
							
						END_IF
				   ELSE
					    _fPos:=stAxis.stNcTOPLC.fActPos-_fEStopPos;
						
						//IF (stAxis.stPLCTONC.eCommand<>E_Command.COMMAND_ABSOLUTEFORK) THEN
						IF (stAxis.stPLCTONC.nRoadID_1=0)THEN 
							IF (_fPos<stAxis.stPLCTONC.fTargetPos)THEN     //03.20
								RETURN;
							END_IF
						ELSE  //非接驳指令
							IF (stAxis.stNcTOPLC.nCuRoadID=stAxis.stPLCTONC.nRoadID_1) THEN 
							   stAxis.stPLCTONC.stStartPosition.nRoadID:=stAxis.stPLCTONC.nRoadID_1;
							   stAxis.stPLCTONC.stEndPosition.nRoadID:=stAxis.stPLCTONC.nRoadID_1;
							   IF (_fPos<stAxis.stPLCTONC.fTargetPos)THEN     //03.20
								   RETURN;
							   END_IF
						    ELSE
							   stAxis.stPLCTONC.stStartPosition.nRoadID:=stAxis.stPLCTONC.nRoadID_2;
							   stAxis.stPLCTONC.stEndPosition.nRoadID:=stAxis.stPLCTONC.nRoadID_2;
							   IF NOT stAxis.stPLCTONC.bRoadDirection  THEN   //正向 
								    IF (_fPos>stAxis.stPLCTONC.fTargetPos)THEN     //03.20
								        RETURN;
							        END_IF
							   ELSE
								   IF (_fPos<stAxis.stPLCTONC.fTargetPos)THEN     //03.20
								        RETURN;
							       END_IF
							   END_IF
						    END_IF
							
						END_IF
				   END_IF
				   
				   //_fTargetVelo:=stAxis.stNcTOPLC.fActVelo;  07.13 
				   //_fVeloStart:=stAxis.stNcTOPLC.fActVelo;
				   IF NOT GVL_MC.bEmStopVMode THEN   //07.13
					   _fTargetVelo:=stAxis.stNcTOPLC.fActVelo;  
				       _fVeloStart:=stAxis.stNcTOPLC.fActVelo;
				   ELSE
					   _fTargetVelo:=_fPtyVelo;  
				       _fVeloStart:=_fPtyVelo;
				   END_IF
				   _fVeloEnd:=0;
				   //_fAcc:=stAxis.stAxisParam.stDynamicDefault.fMaxDeceleration;
				   //_fDec:=stAxis.stAxisParam.stDynamicDefault.fMaxDeceleration;
				   _fAcc:=GVL_MC.nMaxDecRatio*stAxis.stPLCTONC.stEndPosition.fAccleration;  //07.13
				   _fDec:=GVL_MC.nMaxDecRatio*stAxis.stPLCTONC.stEndPosition.fDeceleration; //07.13	
				   _fDistance:=_fEStopPos;
				   _bEnable:=TRUE;
				   _nPathSegment:=1;
				   //stAxis.stAxisStatus.bSynDecActive:=TRUE;
				   stAxis.stAxisStatus.bSynStopping:=TRUE;
		           _bEstopping:=TRUE;  
				 IF GVL_MC.cDebug  THEN
					_sMessage:=FC_StrContact(stAxis,'pPremover PyEstop path ');
					 ADSLOGSTR(ADSLOG_MSGTYPE_HINT, _sMessage, '');
				END_IF
		END_IF
			
ELSE
	IF (_pNextRoadPremover^.stNcTOPLC.nAxisId<>0)AND (stAxis.stAxisStatus.nNcCycleCounter<>0) THEN 
		_fEStopPos:= 0.5*stAxis.stNcTOPLC.fActVelo*stAxis.stNcTOPLC.fActVelo/(GVL_MC.nMaxDecRatio*stAxis.stPLCTONC.stEndPosition.fDeceleration);  //07.13
			IF _fbTonCuPos.Q  AND NOT _bEstopping  THEN   //02.28 增加实际距离检测
				IF (_eDirection=E_Direction.DIRECTION_POSITIVE)THEN
					_fPos:=_fEStopPos+stAxis.stNcTOPLC.fActPos;
					IF (stAxis.stNcTOPLC.fActPos+_fEStopPos)>_fRoad1_Lenth THEN
						stAxis.stPLCTONC.stStartPosition.nRoadID:=stAxis.stPLCTONC.nRoadID_1;
						stAxis.stPLCTONC.stEndPosition.nRoadID:=stAxis.stPLCTONC.nRoadID_2;
                         IF NOT stAxis.stPLCTONC.bRoadDirection  THEN   //正向 
								 IF (_fPos>stAxis.stPLCTONC.fTargetPos)THEN     //03.20
								      RETURN;
							     END_IF
					     ELSE
								 IF (_fPos<stAxis.stPLCTONC.fTargetPos)THEN     //03.20
								        RETURN;
							     END_IF
					     END_IF
						
					ELSE
						stAxis.stPLCTONC.stStartPosition.nRoadID:=stAxis.stPLCTONC.nRoadID_1;
						stAxis.stPLCTONC.stEndPosition.nRoadID:=stAxis.stPLCTONC.nRoadID_1; 
					END_IF
			    ELSE
			        _fPos:=stAxis.stNcTOPLC.fActPos-_fEStopPos;
					IF (stAxis.stNcTOPLC.fActPos-_fStopPos)<0 THEN
						stAxis.stPLCTONC.stStartPosition.nRoadID:=stAxis.stPLCTONC.nRoadID_1;
						stAxis.stPLCTONC.stEndPosition.nRoadID:=stAxis.stPLCTONC.nRoadID_2; 
						IF NOT stAxis.stPLCTONC.bRoadDirection  THEN   //正向 
							IF (_fPos>stAxis.stPLCTONC.fTargetPos)THEN     //03.20
									  RETURN;
							 END_IF
						ELSE
							IF (_fPos<stAxis.stPLCTONC.fTargetPos)THEN     //03.20
									  RETURN;
							END_IF
					    END_IF
						
					ELSE
						stAxis.stPLCTONC.stStartPosition.nRoadID:=stAxis.stPLCTONC.nRoadID_1;
						stAxis.stPLCTONC.stEndPosition.nRoadID:=stAxis.stPLCTONC.nRoadID_1; 
					END_IF
					
			    END_IF 
			    _fDistance:=_fEStopPos;
                 _fAcc:=GVL_MC.nMaxDecRatio*stAxis.stPLCTONC.stEndPosition.fAccleration;  //07.13
				 _fDec:=GVL_MC.nMaxDecRatio*stAxis.stPLCTONC.stEndPosition.fDeceleration; //07.13	
	
				 IF NOT GVL_MC.bEmStopVMode THEN   //07.13
					   _fTargetVelo:=stAxis.stNcTOPLC.fActVelo;  
				       _fVeloStart:=stAxis.stNcTOPLC.fActVelo;
				   ELSE
					   _fTargetVelo:=_fPtyVelo;  
				       _fVeloStart:=_fPtyVelo;
				   END_IF
				_fVeloEnd:=0;
				_bEnable:=TRUE;
				_nPathSegment:=1;
				stAxis.stAxisStatus.bSynStopping:=TRUE;
				_bEstopping:=TRUE;
				IF GVL_MC.cDebug  THEN
					_sMessage:=FC_StrContact(stAxis,'pNextRoadPremover PyEstop path');
					 ADSLOGSTR(ADSLOG_MSGTYPE_HINT, _sMessage, '');
				END_IF
			END_IF
	   // END_IF			  	  
    END_IF
END_IF
END_ACTION

ACTION A_FollowMasterPlanning:
_stPathRef:=stAxis.stAxisStatus.pMaster^.stAxisStatus.stPathRef;
//_fMasterGap:=stAxis.stAxisStatus.pMaster^.stAxisStatus.stPathRef.fGap-stAxis.stAxisStatus.pMaster^.stAxisParam.fClampLength*0.5;
_fMasterGap:=stAxis.stAxisStatus.pMaster^.stAxisStatus.stPathRef.fGap;
IF (stAxis.stAxisStatus.pMaster^.stAxisStatus.stPathRef._nPathSegmentNum=1)THEN
	IF stAxis.stAxisStatus.pMaster^.stAxisStatus.bPositiveDirection THEN 
	   _stPathRef.aExecutablePath[0].fStartPos:=stAxis.stNcTOPLC.fActPos;
	   IF (stAxis.stAxisStatus.pMaster^.stNcTOPLC.fActPos<stAxis.stNcTOPLC.fActPos)THEN
		   _stPathRef.aExecutablePath[0].fEndPos:=stAxis.stAxisStatus.pMaster^.stAxisStatus.stPathRef.aExecutablePath[0].fEndPos+stAxis.stNcTOPLC.fModuloFactor-stAxis.stAxisStatus.stPathRef.fSlaveGap;
	   ELSE
	       _stPathRef.aExecutablePath[0].fEndPos:=stAxis.stAxisStatus.pMaster^.stAxisStatus.stPathRef.aExecutablePath[0].fEndPos-stAxis.stAxisStatus.stPathRef.fSlaveGap;
	   END_IF
	   
	   _stPathRef.aSafePath[0]:=_stPathRef.aExecutablePath[0];
	   //_stPathRef.aSafePath[0].fStartPos:=_stPathRef.aExecutablePath[0].fStartPos-stAxis.stAxisParam.fClampLength*0.5-_fMasterGap;
	   //_stPathRef.aSafePath[0].fEndPos:=_stPathRef.aExecutablePath[0].fEndPos-stAxis.stAxisParam.fClampLength*0.5-_fMasterGap;
	   _stPathRef.aSafePath[0].fStartPos:=_stPathRef.aExecutablePath[0].fStartPos-stAxis.stAxisParam.fClampLength*0.5;
	   _stPathRef.aSafePath[0].fEndPos:=_stPathRef.aExecutablePath[0].fEndPos-stAxis.stAxisParam.fClampLength*0.5;
    ELSE
	   _stPathRef.aExecutablePath[0].fStartPos:=stAxis.stNcTOPLC.fActPos;
	    IF (stAxis.stAxisStatus.pMaster^.stNcTOPLC.fActPos>stAxis.stNcTOPLC.fActPos)THEN
			_stPathRef.aExecutablePath[0].fEndPos:=stAxis.stAxisStatus.pMaster^.stAxisStatus.stPathRef.aExecutablePath[0].fEndPos-stAxis.stNcTOPLC.fModuloFactor+stAxis.stAxisStatus.stPathRef.fSlaveGap;
		ELSE
			_stPathRef.aExecutablePath[0].fEndPos:=stAxis.stAxisStatus.pMaster^.stAxisStatus.stPathRef.aExecutablePath[0].fEndPos+stAxis.stAxisStatus.stPathRef.fSlaveGap;
		END_IF
	   
	   _stPathRef.aSafePath[0]:=_stPathRef.aExecutablePath[0];
	   //_stPathRef.aSafePath[0].fStartPos:=_stPathRef.aExecutablePath[0].fStartPos+stAxis.stAxisParam.fClampLength*0.5+_fMasterGap;
	   //_stPathRef.aSafePath[0].fEndPos:=_stPathRef.aExecutablePath[0].fEndPos+stAxis.stAxisParam.fClampLength*0.5+_fMasterGap;
	   _stPathRef.aSafePath[0].fStartPos:=_stPathRef.aExecutablePath[0].fStartPos+stAxis.stAxisParam.fClampLength*0.5;
	   _stPathRef.aSafePath[0].fEndPos:=_stPathRef.aExecutablePath[0].fEndPos+stAxis.stAxisParam.fClampLength*0.5;
    END_IF
	
	
ELSIF(stAxis.stAxisStatus.pMaster^.stAxisStatus.stPathRef._nPathSegmentNum=2)THEN 
	IF stAxis.stAxisStatus.pMaster^.stAxisStatus.bPositiveDirection THEN 
	   _stPathRef.aExecutablePath[0].fStartPos:=stAxis.stNcTOPLC.fActPos;
	   IF (stAxis.stAxisStatus.pMaster^.stNcTOPLC.fActPos<stAxis.stNcTOPLC.fActPos)THEN
		   _stPathRef.aExecutablePath[0].fEndPos:=stAxis.stAxisStatus.pMaster^.stAxisStatus.stPathRef.aExecutablePath[0].fEndPos+stAxis.stNcTOPLC.fModuloFactor-stAxis.stAxisStatus.stPathRef.fSlaveGap;
	   ELSE
	       _stPathRef.aExecutablePath[0].fEndPos:=stAxis.stAxisStatus.pMaster^.stAxisStatus.stPathRef.aExecutablePath[0].fEndPos-stAxis.stAxisStatus.stPathRef.fSlaveGap;
	   END_IF
	   //_stPathRef.aExecutablePath[0].fEndPos:=stAxis.stAxisStatus.pMaster^.stAxisStatus.stPathRef.aExecutablePath[0].fEndPos-stAxis.stAxisStatus.stPathRef.fSlaveGap;
	   _stPathRef.aExecutablePath[1].fStartPos:=_stPathRef.aExecutablePath[0].fEndPos;
	   
	   IF (stAxis.stAxisStatus.pMaster^.stNcTOPLC.fActPos<stAxis.stNcTOPLC.fActPos)THEN
		   _stPathRef.aExecutablePath[1].fEndPos:=stAxis.stAxisStatus.pMaster^.stAxisStatus.stPathRef.aExecutablePath[1].fEndPos+stAxis.stNcTOPLC.fModuloFactor-stAxis.stAxisStatus.stPathRef.fSlaveGap;
	   ELSE
	       _stPathRef.aExecutablePath[1].fEndPos:=stAxis.stAxisStatus.pMaster^.stAxisStatus.stPathRef.aExecutablePath[1].fEndPos-stAxis.stAxisStatus.stPathRef.fSlaveGap;
	   END_IF
	   //_stPathRef.aExecutablePath[1].fEndPos:=stAxis.stAxisStatus.pMaster^.stAxisStatus.stPathRef.aExecutablePath[1].fEndPos-stAxis.stAxisStatus.stPathRef.fSlaveGap;
	   _stPathRef.aSafePath[0]:=_stPathRef.aExecutablePath[0];
	   //_stPathRef.aSafePath[0].fStartPos:=_stPathRef.aExecutablePath[0].fStartPos-stAxis.stAxisParam.fClampLength*0.5-_fMasterGap;
	   //_stPathRef.aSafePath[0].fEndPos:=_stPathRef.aExecutablePath[0].fEndPos-stAxis.stAxisParam.fClampLength*0.5-_fMasterGap;
	    _stPathRef.aSafePath[0].fStartPos:=_stPathRef.aExecutablePath[0].fStartPos-stAxis.stAxisParam.fClampLength*0.5;
	    _stPathRef.aSafePath[0].fEndPos:=_stPathRef.aExecutablePath[0].fEndPos-stAxis.stAxisParam.fClampLength*0.5;
	   _stPathRef.aSafePath[1]:=_stPathRef.aExecutablePath[1];
	   //_stPathRef.aSafePath[1].fStartPos:=_stPathRef.aExecutablePath[1].fStartPos-stAxis.stAxisParam.fClampLength*0.5-_fMasterGap;
	   //_stPathRef.aSafePath[1].fEndPos:=_stPathRef.aExecutablePath[1].fEndPos-stAxis.stAxisParam.fClampLength*0.5-_fMasterGap;
	   _stPathRef.aSafePath[1].fStartPos:=_stPathRef.aExecutablePath[1].fStartPos-stAxis.stAxisParam.fClampLength*0.5;
	   _stPathRef.aSafePath[1].fEndPos:=_stPathRef.aExecutablePath[1].fEndPos-stAxis.stAxisParam.fClampLength*0.5;
    ELSE
		_stPathRef.aExecutablePath[0].fStartPos:=stAxis.stNcTOPLC.fActPos;
		IF (stAxis.stAxisStatus.pMaster^.stNcTOPLC.fActPos>stAxis.stNcTOPLC.fActPos)THEN
			_stPathRef.aExecutablePath[0].fEndPos:=stAxis.stAxisStatus.pMaster^.stAxisStatus.stPathRef.aExecutablePath[0].fEndPos-stAxis.stNcTOPLC.fModuloFactor+stAxis.stAxisStatus.stPathRef.fSlaveGap;
		ELSE
			_stPathRef.aExecutablePath[0].fEndPos:=stAxis.stAxisStatus.pMaster^.stAxisStatus.stPathRef.aExecutablePath[0].fEndPos+stAxis.stAxisStatus.stPathRef.fSlaveGap;
		END_IF
	   //_stPathRef.aExecutablePath[0].fEndPos:=stAxis.stAxisStatus.pMaster^.stAxisStatus.stPathRef.aExecutablePath[0].fEndPos+stAxis.stAxisStatus.stPathRef.fSlaveGap;
	   _stPathRef.aExecutablePath[1].fStartPos:=_stPathRef.aExecutablePath[0].fEndPos;
	   
	    IF (stAxis.stAxisStatus.pMaster^.stNcTOPLC.fActPos>stAxis.stNcTOPLC.fActPos)THEN
			_stPathRef.aExecutablePath[1].fEndPos:=stAxis.stAxisStatus.pMaster^.stAxisStatus.stPathRef.aExecutablePath[1].fEndPos-stAxis.stNcTOPLC.fModuloFactor+stAxis.stAxisStatus.stPathRef.fSlaveGap;
		ELSE
			_stPathRef.aExecutablePath[1].fEndPos:=stAxis.stAxisStatus.pMaster^.stAxisStatus.stPathRef.aExecutablePath[1].fEndPos+stAxis.stAxisStatus.stPathRef.fSlaveGap;
		END_IF
	   //_stPathRef.aExecutablePath[1].fEndPos:=stAxis.stAxisStatus.pMaster^.stAxisStatus.stPathRef.aExecutablePath[1].fEndPos+stAxis.stAxisStatus.stPathRef.fSlaveGap;
	   _stPathRef.aSafePath[0]:=_stPathRef.aExecutablePath[0];
	   //_stPathRef.aSafePath[0].fStartPos:=_stPathRef.aExecutablePath[0].fStartPos+stAxis.stAxisParam.fClampLength*0.5+_fMasterGap;
	   //_stPathRef.aSafePath[0].fEndPos:=_stPathRef.aExecutablePath[0].fEndPos+stAxis.stAxisParam.fClampLength*0.5+_fMasterGap;
	   _stPathRef.aSafePath[0].fStartPos:=_stPathRef.aExecutablePath[0].fStartPos+stAxis.stAxisParam.fClampLength*0.5;
	   _stPathRef.aSafePath[0].fEndPos:=_stPathRef.aExecutablePath[0].fEndPos+stAxis.stAxisParam.fClampLength*0.5;
	   _stPathRef.aSafePath[1]:=_stPathRef.aExecutablePath[1];
	   //_stPathRef.aSafePath[1].fStartPos:=_stPathRef.aExecutablePath[1].fStartPos+stAxis.stAxisParam.fClampLength*0.5+_fMasterGap;
	   //_stPathRef.aSafePath[1].fEndPos:=_stPathRef.aExecutablePath[1].fEndPos+stAxis.stAxisParam.fClampLength*0.5+_fMasterGap;
	   _stPathRef.aSafePath[1].fStartPos:=_stPathRef.aExecutablePath[1].fStartPos+stAxis.stAxisParam.fClampLength*0.5;
	   _stPathRef.aSafePath[1].fEndPos:=_stPathRef.aExecutablePath[1].fEndPos+stAxis.stAxisParam.fClampLength*0.5;
	END_IF

ELSE
	;
   
END_IF


stAxis.stAxisStatus.stPathRef:=_stPathRef;
//stAxis.stAxisStatus.stPathRef.fGap:=_fMasterGap+stAxis.stAxisParam.fClampLength*0.5;

stAxis.stPLCTONC.fTargetVelocity:=stAxis.stAxisStatus.pMaster^.stPLCTONC.fTargetVelocity;
IF stAxis.stAxisStatus.pMaster^.stPLCTONC.bCmdDceUpdate THEN
   stAxis.stAxisStatus.bSynDecActive:=TRUE;
END_IF
_fTime:=0;
_nIndex:=0;
stAxis.stAxisStatus.nNcCycleCounter:=0;
stAxis.stAxisStatus.stPathRef.bCalculateDone:=TRUE;
_bCalculateDone:=TRUE;
END_ACTION

ACTION A_FollowMaterPosition:
_nSysType:=stAxis.stPLCTONC.nSysType;
stAxis.stNcTOPLC.nAxisState:=6;  //03.14
stAxis.stAxisStatus.nNcCycleCounter:=stAxis.stAxisStatus.pMaster^.stAxisStatus.nNcCycleCounter;
//stAxis.stNcTOPLC.fSetVelo:=floor(stAxis.stAxisStatus.pMaster^.stNcTOPLC.fActVelo*stAxis.stPLCTONC.fGearRatio);  //04.15注释
stAxis.stNcTOPLC.fActVelo:=LTRUNC(stAxis.stAxisStatus.pMaster^.stNcTOPLC.fActVelo*stAxis.stPLCTONC.fGearRatio);
IF (_eDirection=E_Direction.DIRECTION_POSITIVE)THEN    //04.15速度方向处理
	  stAxis.stNcTOPLC.fSetVelo:=stAxis.stNcTOPLC.fActVelo;
ELSE
      stAxis.stNcTOPLC.fSetVelo:=-stAxis.stNcTOPLC.fActVelo;
END_IF

(*IF stAxis.stAxisStatus.bPositiveDirection THEN
    stAxis.stNcTOPLC.fActPos:=stAxis.stAxisStatus.pMaster^.stNcTOPLC.fDealtPos*stAxis.stPLCTONC.fGearRatio +stAxis.stNcTOPLC.fActPos;

ELSE
    stAxis.stNcTOPLC.fActPos:=-stAxis.stAxisStatus.pMaster^.stNcTOPLC.fDealtPos*stAxis.stPLCTONC.fGearRatio +stAxis.stNcTOPLC.fActPos;
END_IF*)

IF (stAxis.stAxisStatus.nNcCycleCounter=0)THEN 
	_stAxis_Point.fPosition:=stAxis.stNcTOPLC.fActPos;
	RETURN;
END_IF
IF stAxis.stAxisStatus.bPositiveDirection THEN
    _stAxis_Point.fPosition:=stAxis.stAxisStatus.pMaster^.stNcTOPLC.fDealtPos*stAxis.stPLCTONC.fGearRatio +_stAxis_Point.fPosition;

ELSE
    _stAxis_Point.fPosition:=-stAxis.stAxisStatus.pMaster^.stNcTOPLC.fDealtPos*stAxis.stPLCTONC.fGearRatio +_stAxis_Point.fPosition;
END_IF
_fRoad1_Lenth:=stAxis.stAxisStatus.pMaster^.stPLCTONC.fRoad1_Length;
_fRoad2_Lenth:=stAxis.stAxisStatus.pMaster^.stPLCTONC.fRoad2_Length;

//  实时位置、速度处理
IF (_nSysType=1)OR(_nSysType=4)	THEN    //接驳线和分叉线
	IF (_eDirection=E_Direction.DIRECTION_POSITIVE)THEN
		IF (stAxis.stAxisStatus.pMaster^.stPLCTONC.nRoadID_1<>0)AND (stAxis.stAxisStatus.pMaster^.stPLCTONC.nRoadID_2<>0)THEN    //id不相同处理
			IF (_stAxis_Point.fPosition<=_fRoad1_Lenth)THEN
				stAxis.stNcTOPLC.fActPos:=_stAxis_Point.fPosition;
				stAxis.stNcTOPLC.nCuRoadID:=stAxis.stAxisStatus.pMaster^.stPLCTONC.nRoadID_1;
			ELSE
				IF NOT stAxis.stAxisStatus.pMaster^.stPLCTONC.bRoadDirection THEN 
				   stAxis.stNcTOPLC.fActPos:=FC_TransformPosition(fOffset:=-_fRoad1_Lenth , fPosition:=_stAxis_Point.fPosition );

				ELSE
					_fPosTemp:=FC_TransformPosition(fOffset:=-_fRoad1_Lenth , fPosition:=_stAxis_Point.fPosition );
					stAxis.stNcTOPLC.fActPos:= _fRoad2_Lenth-_fPosTemp;
				END_IF
				
				stAxis.stNcTOPLC.nCuRoadID:=stAxis.stAxisStatus.pMaster^.stPLCTONC.nRoadID_2;
			END_IF
		
		END_IF
	ELSE
		
		IF (stAxis.stAxisStatus.pMaster^.stPLCTONC.nRoadID_1<>0)AND (stAxis.stAxisStatus.pMaster^.stPLCTONC.nRoadID_2<>0)THEN    //id不相同处理   //id不相同处理
			IF (_stAxis_Point.fPosition>=0)THEN
				stAxis.stNcTOPLC.nCuRoadID:=stAxis.stAxisStatus.pMaster^.stPLCTONC.nRoadID_1;
				stAxis.stNcTOPLC.fActPos:=_stAxis_Point.fPosition;
				
			ELSE
				IF NOT stAxis.stAxisStatus.pMaster^.stPLCTONC.bRoadDirection THEN     //正向
					stAxis.stNcTOPLC.fActPos:=ABS(_stAxis_Point.fPosition);
				ELSE
					_fPosTemp:=ABS(_stAxis_Point.fPosition);
					stAxis.stNcTOPLC.fActPos:= _fRoad2_Lenth-_fPosTemp;
				END_IF
				
				stAxis.stNcTOPLC.nCuRoadID:=stAxis.stAxisStatus.pMaster^.stPLCTONC.nRoadID_2;
			END_IF
              
		END_IF
	
	END_IF
	
ELSE
    stAxis.stNcTOPLC.fDealtPos:=ABS(LTRUNC(_stAxis_Point.fPosition)-stAxis.stNcTOPLC.fActPos);    //01.13
	stAxis.stNcTOPLC.fActPos:=LTRUNC(_stAxis_Point.fPosition);
  
END_IF
END_ACTION

ACTION A_FollowPlanning:
_fMasterEndPos:=0;
//_fMasterStartPos:=0;

_fMasterStartPos:=stAxis.stAxisStatus.pMaster^.stNcTOPLC.fActPos;

_bCalculateDone:=TRUE;
END_ACTION

ACTION A_FollowPosition:
stAxis.stAxisStatus.nNcCycleCounter:=stAxis.stAxisStatus.nNcCycleCounter+1;
_fMasterEndPos:=stAxis.stAxisStatus.pMaster^.stNcTOPLC.fActPos;

_fDePos:=_fMasterEndPos-_fMasterStartPos;
_fVeloRatio:=stAxis.stPLCTONC.fGearRatio;
//_fVeloRatio:=stAxis.stAxisStatus.stPathRef.fVeloRatio;
//stAxis.stNcTOPLC.fSetPos:=stAxis.stNcTOPLC.fActPos+_fVeloRatio*_fDePos;
stAxis.stNcTOPLC.fActPos:=stAxis.stNcTOPLC.fActPos+_fVeloRatio*_fDePos;
stAxis.stNcTOPLC.fSetVelo:=stAxis.stAxisStatus.pMaster^.stNcTOPLC.fActVelo*_fVeloRatio;
//stAxis.stNcTOPLC.fSetVelo:=_fDePos/fCycleTime;

IF (_fDePos=0) THEN
	
	stAxis.stNcTOPLC.fSetVelo:=stAxis.stNcTOPLC.fActVelo;
END_IF

//stAxis.stNcTOPLC.fActPos:=stAxis.stNcTOPLC.fSetPos;
stAxis.stNcTOPLC.fActVelo:=stAxis.stNcTOPLC.fSetVelo;

(*IF stAxis.stAxisStatus.bPositiveDirection THEN
	stAxis.stNcTOPLC.nModuloSetTurns:=LREAL_TO_DINT(LTRUNC(stAxis.stNcTOPLC.fSetPos/stAxis.stNcTOPLC.fModuloFactor));
ELSE
	IF stAxis.stNcTOPLC.fSetPos<(stAxis.stNcTOPLC.nModuloSetTurns*stAxis.stNcTOPLC.fModuloFactor)THEN 
			stAxis.stNcTOPLC.nModuloSetTurns:=stAxis.stNcTOPLC.nModuloSetTurns-1;
	END_IF
END_IF

stAxis.stNcTOPLC.fModuloSetPos:= MODABS(stAxis.stNcTOPLC.fSetPos,stAxis.stNcTOPLC.fModuloFactor);*)

_fMasterStartPos:=stAxis.stAxisStatus.pMaster^.stNcTOPLC.fActPos;
END_ACTION

ACTION A_GapControl:

(*****
   1. 判断前后动子距离优先触发减速
   2. 如果前后距离与防碰撞距离小于一定阈值优先触发同步减速功能
   3. 如果是前动子自动触发减速，会出现后动子先减速到目标速度，前动子后减速到目标速度,前后动子距离会变大一点
****)
_fbDecPathTrig(CLK:=_pPremover^.stPLCTONC.bCmdDceUpdate OR _pPremover^.stAxisStatus.bSynDecActive  , Q=> );// 同步时前动子减速  03.28注释
IF (_pPremover^.stAxisStatus.nNcCycleCounter<>0)THEN 
	 A_CatchUp();
	//IF ((_fRealDis -_fGapSet)<=cDealtGap) THEN    //10.18 
	  IF ((_fRealDis -_fGapSet)<=_fSetDealtGap) THEN  
		IF _fbDecPathTrig.Q THEN 
		   // 04.02 增加road2情况
		   IF (stAxis.stPLCTONC.nRoadID_2<>0)AND (stAxis.stPLCTONC.nRoadID_1<>0)AND(stAxis.stNcTOPLC.nCuRoadID=stAxis.stPLCTONC.nRoadID_2)THEN
			   IF (stAxis.stPLCTONC.stStartPosition.nRoadID<>stAxis.stPLCTONC.stEndPosition.nRoadID)THEN
					IF (_eDirection=E_Direction.DIRECTION_POSITIVE)THEN
						IF NOT stAxis.stPLCTONC.bRoadDirection  THEN
							 _fPos:=stAxis.stPLCTONC.stEndPosition.fPosition-stAxis.stPLCTONC.fRoad1_Length;
						ELSE
							_fPos:=stAxis.stPLCTONC.fRoad2_Length-(stAxis.stPLCTONC.stEndPosition.fPosition-stAxis.stPLCTONC.fRoad1_Length);
						END_IF
						_fDistance:=ABS(stAxis.stNcTOPLC.fActPos-_fPos);
					ELSE
						IF NOT stAxis.stPLCTONC.bRoadDirection  THEN
							 _fPos:=ABS(stAxis.stPLCTONC.stEndPosition.fPosition);
						ELSE
							_fPos:=stAxis.stPLCTONC.fRoad2_Length-ABS(stAxis.stPLCTONC.stEndPosition.fPosition);
						END_IF
						_fDistance:=ABS(stAxis.stNcTOPLC.fActPos-_fPos);
					END_IF
			   ELSE
					_fPos:=stAxis.stPLCTONC.stEndPosition.fPosition;
					_fDistance:=ABS(stAxis.stNcTOPLC.fActPos-_fPos);
			   END_IF
		   ELSE
			   _fPos:=stAxis.stPLCTONC.stEndPosition.fPosition;
			   IF (_eDirection=E_Direction.DIRECTION_POSITIVE)THEN
				  _fDistance:=_fPos-stAxis.stNcTOPLC.fActPos;
			   ELSE
				  _fDistance:=stAxis.stNcTOPLC.fActPos-_fPos;
			   END_IF
		   END_IF
		   //_fPos:=stAxis.stPLCTONC.stEndPosition.fPosition;
		   _fTargetVelo:=_pPremover^.stAxisStatus.stPathRef.fTargetVelocity;
		   _fVeloStart:=stAxis.stNcTOPLC.fActVelo;
		   _fVeloEnd:=0;
		   _fAcc:=stAxis.stPLCTONC.stEndPosition.fAccleration;
		   _fDec:=stAxis.stPLCTONC.stEndPosition.fDeceleration;
		   
		   _bEnable:=TRUE;
		   _nPathSegment:=1;
		   stAxis.stAxisStatus.bSynDecActive:=TRUE;
		   IF GVL_MC.cDebug  THEN
			_sMessage:=FC_StrContact(stAxis,'SynDecActive path');
			 ADSLOGSTR(ADSLOG_MSGTYPE_HINT, _sMessage, '');
		   END_IF
		END_IF
	 END_IF
END_IF

//模式控制
END_ACTION

ACTION A_GetPosition:
IF (stAxis.stPLCTONC.ePlanningMode=E_PlanningMode.PLANNINGMODE_TSHAPED)THEN 
   A_TShapedPosition();
   _bEndOfProfile:=FALSE;
ELSIF (stAxis.stPLCTONC.ePlanningMode=E_PlanningMode.PLANNINGMODE_SSHAPED)THEN 
  A_SShapedPosition();
ELSIF (stAxis.stPLCTONC.ePlanningMode=E_PlanningMode.PLANNINGMODE_LINEAR)THEN 
  A_LinearPosition();
 
ELSIF (stAxis.stPLCTONC.ePlanningMode=E_PlanningMode.PLANNINGMODE_FOLLOWMASTER)THEN 
	//A_TShapedPosition();
    A_FollowMaterPosition();
ELSIF (stAxis.stPLCTONC.ePlanningMode=E_PlanningMode.PLANNINGMODE_PLOYNOM3)THEN 
	A_Ploynom3Position();
ELSIF (stAxis.stPLCTONC.ePlanningMode=E_PlanningMode.PLANNINGMODE_PLOYNOM5)THEN
    IF NOT _bEndOfProfile THEN 
	    A_Ploynom5Position();
    ELSE           //12.31
        A_ContantVeloPosition();
    END_IF 	
ELSIF (stAxis.stPLCTONC.ePlanningMode=E_PlanningMode.PLANNINGMODE_FOLLOW)THEN 
	A_FollowPosition();	
ELSE 
    A_TShapedPosition();
    _bEndOfProfile:=FALSE;
END_IF
END_ACTION

ACTION A_LinearPlanning:
_nIndex:=1;
stAxis.stAxisStatus.nNcCycleCounter:=0;
IF (stAxis.stPLCTONC.nLinearPointNum<>0)THEN 
   _fLinearDealt:=(_fPos-stAxis.stNcTOPLC.fActPos)/stAxis.stPLCTONC.nLinearPointNum;
END_IF 

FOR  _nPointIndex:=1 TO stAxis.stPLCTONC.nLinearPointNum  DO
	_aLinearPosition[_nPointIndex]:=stAxis.stNcTOPLC.fActPos+_fLinearDealt*_nPointIndex;
END_FOR

_bCalculateDone:=TRUE;
END_ACTION

ACTION A_LinearPosition:

stAxis.stNcTOPLC.fActPos:=_aLinearPosition[_nIndex];

stAxis.stNcTOPLC.fSetVelo:=stAxis.stPLCTONC.stEndPosition.fVelocity;
stAxis.stNcTOPLC.fActVelo:=stAxis.stPLCTONC.stEndPosition.fVelocity;
_nIndex:=_nIndex+1;
IF (_aLinearPosition[_nIndex]=0)THEN 
	 _bCalculateDone:=FALSE;
	 _nIndex:=0;
END_IF

IF (_nIndex>UINT_TO_INT(stAxis.stPLCTONC.nLinearPointNum))THEN 
	_bCalculateDone:=FALSE;
	_nIndex:=0;
END_IF
END_ACTION

ACTION A_NCStartCase:
//根据不同指令控制NC路径规划 
// 命令触发
_fbTrig(CLK:=stAxis.stPLCTONC.bNcStart , Q=> );
IF _fbTrig.Q  THEN 
	_nPathSegment:=1;
	_fPos:=stAxis.stPLCTONC.stEndPosition.fPosition;
	_fStartPos:=stAxis.stNcTOPLC.fActPos;
	_fEndPos:=stAxis.stPLCTONC.stEndPosition.fPosition;
	_fTargetVelo:=stAxis.stPLCTONC.fTargetVelocity;
	
	IF (stAxis.stAxisStatus.nNcCycleCounter=0)THEN
		_fVeloStart:=0;  
		//_fVeloEnd:=0;   //12.03
		_fVeloEnd:=stAxis.stPLCTONC.stEndPosition.fVelocity;  //12.03
	ELSE
	    _fVeloStart:=stAxis.stNcTOPLC.fActVelo;
		//_fVeloEnd:=0;  //12.03
		_fVeloEnd:=stAxis.stPLCTONC.stEndPosition.fVelocity;  //12.03
	END_IF
	IF stAxis.stAxisStatus.bSlave THEN
		_fVeloStart:=stAxis.stNcTOPLC.fActVelo;
		_fVeloEnd:=0;
	END_IF
	
	IF (_eDirection=E_Direction.DIRECTION_POSITIVE)THEN
	     _fDistance:=_fPos-stAxis.stNcTOPLC.fActPos;
    ELSE
        _fDistance:=stAxis.stNcTOPLC.fActPos-_fPos;
    END_IF 
	// 04.08
	IF (stAxis.stPLCTONC.nRoadID_1<>0) AND (stAxis.stPLCTONC.nRoadID_2<>0)THEN
		IF (stAxis.stPLCTONC.stStartPosition.nRoadID=stAxis.stPLCTONC.nRoadID_2)THEN
			IF NOT stAxis.stPLCTONC.bRoadDirection  THEN   //正向 
                 _fDistance:=_fPos-stAxis.stNcTOPLC.fActPos;
            ELSE
                 _fDistance:=stAxis.stNcTOPLC.fActPos-_fPos;
            END_IF 
		END_IF
	END_IF
	// 04.08
	IF (stAxis.stPLCTONC.ePlanningMode<>E_PlanningMode.PLANNINGMODE_LINEAR)AND (stAxis.stPLCTONC.ePlanningMode<>E_PlanningMode.PLANNINGMODE_FOLLOW)THEN 
		IF (_fDistance<=0) AND (stAxis.stPLCTONC.ePlanningMode=E_PlanningMode.PLANNINGMODE_TSHAPED)  THEN 
			RETURN ;
		END_IF
	END_IF 
	_fAcc:=stAxis.stPLCTONC.stEndPosition.fAccleration;
	_fDec:=stAxis.stPLCTONC.stEndPosition.fDeceleration;
	_fJerk:=stAxis.stPLCTONC.stEndPosition.fbJerk;
	_fGap:=stAxis.stAxisStatus.stPathRef.fGap;
	_bEnable:=TRUE;
	_bSynMode:=FALSE;
	//_pPremover^.stAxisStatus.bSynDecActive:=FALSE;

	IF GVL_MC.cDebug  THEN
		_sMessage:=FC_StrContact(stAxis,'NC generate path');
	     ADSLOGSTR(ADSLOG_MSGTYPE_HINT, _sMessage, '');	 
    END_IF
	 _nSysType:=stAxis.stPLCTONC.nSysType;    //01.13
	 
	 IF stAxis.stAxisStatus.bStoppingFlag THEN    //10.09 注释
		  stAxis.stAxisStatus.bSynStopping:=TRUE;
	 END_IF
	
	 
END_IF
IF (stAxis.stAxisStatus.pMaster<>0)THEN 
   _fbSlaveTrig(CLK:=(stAxis.stAxisStatus.pMaster^.stPLCTONC.bNcStart OR stAxis.stAxisStatus.pMaster^.stAxisStatus.bSynDecActive)
          AND stAxis.stAxisStatus.pMaster^.stAxisStatus.stPathRef.bCalculateDone  , Q=> );
END_IF 
IF (stAxis.stPLCTONC.eCommand=E_Command.COMMAND_ABSOLUTE)OR (stAxis.stPLCTONC.eCommand=E_Command.COMMAND_ABSOLUTEFORK)THEN 
		
   IF (_pPremover^.stAxisStatus.nNcCycleCounter<>0) AND (stAxis.stAxisStatus.nNcCycleCounter<>0)AND NOT stAxis.stAxisStatus.bSynStopping THEN 
	
		IF (_pPremover^.stAxisStatus.stPathRef.fTargetVelocity <>stAxis.stAxisStatus.stPathRef.fTargetVelocity) THEN
			   A_GapControl();
		END_IF
   ELSE     //03.18  增加下一段road处理
		 IF (_pNextRoadPremover^.stAxisStatus.nNcCycleCounter<>0)AND (stAxis.stAxisStatus.nNcCycleCounter<>0)AND NOT stAxis.stAxisStatus.bSynStopping    
			AND(_pNextRoadPremover^.stAxisStatus.stPathRef.fTargetVelocity <>stAxis.stAxisStatus.stPathRef.fTargetVelocity) THEN   //10.28
			  A_NextRoadGapControl(); 
		  END_IF
	   
   END_IF
	
   _fbPathTrig(CLK:= _pPremover^.stAxisStatus.bSynDecActive, Q=> );  //重新触发gap调节
   IF _fbPathTrig.Q THEN 
	   _bSynMode:=FALSE;
   END_IF
	   
ELSIF (stAxis.stPLCTONC.eCommand=E_Command.COMMAND_GEARIN)OR(stAxis.stPLCTONC.eCommand=E_Command.COMMAND_CAMIN)THEN 
	   IF _fbSlaveTrig.Q THEN
	//	   _bEnable:=TRUE;
	            ;
	   END_IF
	   _bCalculateDone:=TRUE;
	   
ELSE 
		; 
END_IF 


 _fbTon(IN:=stAxis.stAxisStatus.bSynDecActive , PT:=T#20MS , Q=> , ET=> );
IF _fbTon.Q THEN
	stAxis.stAxisStatus.bSynDecActive:=FALSE;
 END_IF
 

// 急停及同步停止处理
IF NOT stAxis.stAxisStatus.bStoppingFlag THEN 	  //03.12 
  A_StopHandle(); 
 
END_IF
END_ACTION

ACTION A_NextPathUpdateNewTarPos:
_fAcc:=stAxis.stPLCTONC.stEndPosition.fAccleration;
_fDec:=stAxis.stPLCTONC.stEndPosition.fDeceleration;
//根据下一段road指令分类

IF (_pNextRoadPremover^.stPLCTONC.nRoadID_1<>0)THEN     //fork指令
	IF (_pNextRoadPremover^.stPLCTONC.stStartPosition.nRoadID<>_pNextRoadPremover^.stPLCTONC.stEndPosition.nRoadID)THEN
		IF (_pNextRoadPremover^.stPLCTONC.stStartPosition.nRoadID=stAxis.stPLCTONC.stStartPosition.nRoadID)THEN  //起点road相同
			IF (_eDirection=E_Direction.DIRECTION_POSITIVE)THEN
				_fUpNewPos:=_pNextRoadPremover^.stAxisStatus.stPathRef.aExecutablePath[0].fEndPos-_fGapSet-stAxis.stNcTOPLC.fActPos;
			ELSE
				_fUpNewPos:=stAxis.stNcTOPLC.fActPos-_pNextRoadPremover^.stAxisStatus.stPathRef.aExecutablePath[0].fEndPos-_fGapSet;
			END_IF
			stAxis.stPLCTONC.stStartPosition.nRoadID:=stAxis.stNcTOPLC.nCuRoadID;
			IF (stAxis.stNcTOPLC.fActPos+_fUpNewPos)>stAxis.stPLCTONC.fRoad1_Length THEN
				 
				 stAxis.stPLCTONC.stEndPosition.nRoadID:=stAxis.stPLCTONC.nRoadID_2;
			ELSE
				 stAxis.stPLCTONC.stEndPosition.nRoadID:=stAxis.stNcTOPLC.nCuRoadID;
			END_IF
		ELSE
			IF (_eDirection=E_Direction.DIRECTION_POSITIVE)THEN
				IF NOT stAxis.stPLCTONC.bRoadDirection  THEN  //正向
				    _fUpNewPos:=_pNextRoadPremover^.stAxisStatus.stPathRef.aExecutablePath[0].fEndPos+stAxis.stPLCTONC.fRoad1_Length-_fGapSet-stAxis.stNcTOPLC.fActPos;
				ELSE
					_fUpNewPos:=stAxis.stPLCTONC.fRoad2_Length-_pNextRoadPremover^.stAxisStatus.stPathRef.aExecutablePath[0].fEndPos+stAxis.stPLCTONC.fRoad1_Length-_fGapSet-stAxis.stNcTOPLC.fActPos;
				END_IF
				IF (stAxis.stNcTOPLC.fActPos+_fUpNewPos)>stAxis.stPLCTONC.fRoad1_Length THEN
				 
					 stAxis.stPLCTONC.stEndPosition.nRoadID:=stAxis.stPLCTONC.nRoadID_2;
				ELSE
					 stAxis.stPLCTONC.stEndPosition.nRoadID:=stAxis.stNcTOPLC.nCuRoadID;
				END_IF
			ELSE
				IF NOT stAxis.stPLCTONC.bRoadDirection  THEN  //正向
				    _fUpNewPos:=stAxis.stNcTOPLC.fActPos+_pNextRoadPremover^.stAxisStatus.stPathRef.aExecutablePath[0].fEndPos-_fGapSet;
				ELSE
					_fUpNewPos:=stAxis.stNcTOPLC.fActPos+_pNextRoadPremover^.stAxisStatus.stPathRef.aExecutablePath[0].fEndPos-stAxis.stPLCTONC.fRoad2_Length-_fGapSet;
				END_IF
				IF (stAxis.stNcTOPLC.fActPos-_fUpNewPos)<0 THEN
			 
					 stAxis.stPLCTONC.stEndPosition.nRoadID:=stAxis.stPLCTONC.nRoadID_2;
				ELSE
					 stAxis.stPLCTONC.stEndPosition.nRoadID:=stAxis.stNcTOPLC.nCuRoadID;
				END_IF
			END_IF
			
		END_IF
	ELSE   //fork指令 根据前动子的edpos id 和当前动子roadid分类讨论
		
		IF (_eDirection=E_Direction.DIRECTION_POSITIVE)THEN
				IF NOT stAxis.stPLCTONC.bRoadDirection  THEN  //正向
				    _fUpNewPos:=_pNextRoadPremover^.stAxisStatus.stPathRef.aExecutablePath[0].fEndPos+stAxis.stPLCTONC.fRoad1_Length-_fGapSet-stAxis.stNcTOPLC.fActPos;
				ELSE
					_fUpNewPos:=stAxis.stPLCTONC.fRoad2_Length-_pNextRoadPremover^.stAxisStatus.stPathRef.aExecutablePath[0].fEndPos+stAxis.stPLCTONC.fRoad1_Length-_fGapSet-stAxis.stNcTOPLC.fActPos;
				END_IF
				stAxis.stPLCTONC.stStartPosition.nRoadID:=stAxis.stNcTOPLC.nCuRoadID;
				IF (stAxis.stNcTOPLC.fActPos+_fUpNewPos)>stAxis.stPLCTONC.fRoad1_Length THEN
					 
					 stAxis.stPLCTONC.stEndPosition.nRoadID:=stAxis.stPLCTONC.nRoadID_2;
				ELSE
					 stAxis.stPLCTONC.stEndPosition.nRoadID:=stAxis.stNcTOPLC.nCuRoadID;
				END_IF
				
		ELSE
				IF NOT stAxis.stPLCTONC.bRoadDirection  THEN  //正向
				    _fUpNewPos:=stAxis.stNcTOPLC.fActPos+_pNextRoadPremover^.stAxisStatus.stPathRef.aExecutablePath[0].fEndPos-_fGapSet;
				ELSE
					//_fUpNewPos:=stAxis.stNcTOPLC.fActPos+_pNextRoadPremover^.stAxisStatus.stPathRef.aExecutablePath[0].fEndPos-stAxis.stPLCTONC.fRoad2_Length-_fGapSet;
					_fUpNewPos:=stAxis.stNcTOPLC.fActPos-_pNextRoadPremover^.stAxisStatus.stPathRef.aExecutablePath[0].fEndPos+stAxis.stPLCTONC.fRoad2_Length-_fGapSet;  //08.20
				END_IF
				stAxis.stPLCTONC.stStartPosition.nRoadID:=stAxis.stNcTOPLC.nCuRoadID;
				IF (stAxis.stNcTOPLC.fActPos-_fUpNewPos)<0 THEN
					 
					 stAxis.stPLCTONC.stEndPosition.nRoadID:=stAxis.stPLCTONC.nRoadID_2;
				ELSE
					 stAxis.stPLCTONC.stEndPosition.nRoadID:=stAxis.stNcTOPLC.nCuRoadID;
				END_IF
				
		END_IF
		 //stAxis.stPLCTONC.stStartPosition.nRoadID:=stAxis.stNcTOPLC.nCuRoadID;
		// stAxis.stPLCTONC.stEndPosition.nRoadID:=stAxis.stNcTOPLC.nCuRoadID;
	END_IF
ELSE   //非fork指令
	IF (_eDirection=E_Direction.DIRECTION_POSITIVE)THEN
		IF NOT stAxis.stPLCTONC.bRoadDirection  THEN  //正向
		   _fUpNewPos:=_pNextRoadPremover^.stAxisStatus.stPathRef.aExecutablePath[0].fEndPos+stAxis.stPLCTONC.fRoad1_Length-_fGapSet-stAxis.stNcTOPLC.fActPos;
	    ELSE
			_fUpNewPos:=stAxis.stPLCTONC.fRoad2_Length-_pNextRoadPremover^.stAxisStatus.stPathRef.aExecutablePath[0].fEndPos+stAxis.stPLCTONC.fRoad1_Length-_fGapSet-stAxis.stNcTOPLC.fActPos;
		END_IF
		stAxis.stPLCTONC.stStartPosition.nRoadID:=stAxis.stNcTOPLC.nCuRoadID;
		IF (stAxis.stNcTOPLC.fActPos+_fUpNewPos)>stAxis.stPLCTONC.fRoad1_Length THEN
			 
		     stAxis.stPLCTONC.stEndPosition.nRoadID:=stAxis.stPLCTONC.nRoadID_2;
		ELSE
			 stAxis.stPLCTONC.stEndPosition.nRoadID:=stAxis.stNcTOPLC.nCuRoadID;
		END_IF
	ELSE
		IF NOT stAxis.stPLCTONC.bRoadDirection  THEN  //正向
			_fUpNewPos:=stAxis.stNcTOPLC.fActPos+_pNextRoadPremover^.stAxisStatus.stPathRef.aExecutablePath[0].fEndPos-_fGapSet;
		ELSE
			//_fUpNewPos:=stAxis.stNcTOPLC.fActPos+_pPremover^.stAxisStatus.stPathRef.aExecutablePath[0].fEndPos-stAxis.stPLCTONC.fRoad2_Length-_fGapSet;
			_fUpNewPos:=stAxis.stNcTOPLC.fActPos-_pNextRoadPremover^.stAxisStatus.stPathRef.aExecutablePath[0].fEndPos+stAxis.stPLCTONC.fRoad2_Length-_fGapSet;  //08.20
		END_IF
        stAxis.stPLCTONC.stStartPosition.nRoadID:=stAxis.stNcTOPLC.nCuRoadID;
		IF (stAxis.stNcTOPLC.fActPos-_fUpNewPos)<0 THEN
			 
		     stAxis.stPLCTONC.stEndPosition.nRoadID:=stAxis.stPLCTONC.nRoadID_2;
		ELSE
			 stAxis.stPLCTONC.stEndPosition.nRoadID:=stAxis.stNcTOPLC.nCuRoadID;
		END_IF	
	END_IF
END_IF
	
_fDistance:=_fUpNewPos;
// 11.01 停止计算距离，根据距离设置目标速度
IF _fDec<>0 THEN  //11.01 
   _fLastPosDeat:=0.5*stAxis.stNcTOPLC.fActVelo*stAxis.stNcTOPLC.fActVelo/_fDec;
END_IF 
IF LTRUNC(_fDistance)<=_fLastPosDeat THEN
	_fTargetVelo:=stAxis.stNcTOPLC.fActVelo;
ELSE
	_fTargetVelo:=stAxis.stPLCTONC.fTargetVelocity;
END_IF

//_fTargetVelo:=stAxis.stNcTOPLC.fActVelo;
_fVeloStart:=stAxis.stNcTOPLC.fActVelo;
_fVeloEnd:=0;
_bEnable:=TRUE;
_nPathSegment:=1;
stAxis.stAxisStatus.bSynStopping:=TRUE;  //10.28

IF GVL_MC.cDebug  THEN
	_sMessage:=FC_StrContact(stAxis,'SynStoping Nextpath');
	 ADSLOGSTR(ADSLOG_MSGTYPE_HINT, _sMessage, '');
END_IF
END_ACTION

ACTION A_NextRoadAccSegmengt:

_fPreTaVel:=_pNextRoadPremover^.stAxisStatus.stPathRef.fTargetVelocity;
_fPreCuVel:=_pNextRoadPremover^.stNcTOPLC.fActVelo;
_fPreAcc:=_pNextRoadPremover^.stAxisStatus.stPathRef.aExecutablePath[0].fAccleration;   //有问题

_fCuVel:=stAxis.stNcTOPLC.fActVelo;

IF (_fCuVel>_fPreTaVel)THEN   //速度>前动子目标速度
	    _fDealt_S1:=0.5*(_fPreTaVel-_fPreCuVel)*(_fPreTaVel-_fPreCuVel)/_fAcc;	
		
        IF (_fDealt_S>_fDealt_S1)THEN	   
	         _fNewAcc:=(_fCuVel-_fPreTaVel)*(_fCuVel-_fPreTaVel)*0.5/(_fDealt_S-_fDealt_S1);
			 IF (_fNewAcc>stAxis.stAxisParam.stDynamicDefault.fMaxDeceleration)THEN 
			    _fNewAcc:=stAxis.stAxisParam.stDynamicDefault.fMaxDeceleration;
		     END_IF
		ELSE
			_fNewAcc:=stAxis.stAxisParam.stDynamicDefault.fMaxDeceleration;
		END_IF
		
	    _fDecTime:=	(_fCuVel-_fPreTaVel)/_fNewAcc;
	    _fNewAccDis:=(_fCuVel*_fCuVel-_fPreTaVel*_fPreTaVel)*0.5/_fNewAcc;   //减速面积
	    _fMinDis:=_fPreTaVel*_fPreTaVel*0.5/_fAcc+_fNewAccDis;  //减速面积+停止最小面积
	    _fPos:=stAxis.stPLCTONC.stEndPosition.fPosition;
	    IF(_fReminDis< _fMinDis)THEN
			_fVeloStart:=stAxis.stNcTOPLC.fActVelo;
			_fVeloEnd:=0.0;
			_fTargetVelo:=_pNextRoadPremover^.stAxisStatus.stPathRef.fTargetVelocity;
			_fAcc:=stAxis.stPLCTONC.stEndPosition.fAccleration;
			_fDec:=stAxis.stPLCTONC.stEndPosition.fDeceleration;
			IF (stAxis.stPLCTONC.nRoadID_2<>0)AND (stAxis.stPLCTONC.nRoadID_1<>0)THEN   //判断指令
				IF (stAxis.stPLCTONC.stStartPosition.nRoadID<>stAxis.stPLCTONC.stEndPosition.nRoadID)THEN
				    IF(stAxis.stNcTOPLC.nCuRoadID=stAxis.stPLCTONC.nRoadID_2) THEN //第二路段
						IF (_eDirection=E_Direction.DIRECTION_POSITIVE)THEN
							 IF NOT stAxis.stPLCTONC.bRoadDirection  THEN   //正向 
								 _fDistance:=_fPos-stAxis.stPLCTONC.fRoad1_Length-stAxis.stNcTOPLC.fActPos;
							 ELSE
								 _fDistance:=stAxis.stNcTOPLC.fActPos-(stAxis.stPLCTONC.fRoad2_Length-_fPos+stAxis.stPLCTONC.fRoad1_Length);
							 END_IF
						ELSE
							IF NOT stAxis.stPLCTONC.bRoadDirection  THEN   //正向 
								 _fDistance:=ABS(_fPos)-stAxis.stNcTOPLC.fActPos;
							 ELSE
								 _fDistance:=stAxis.stNcTOPLC.fActPos-(stAxis.stPLCTONC.fRoad2_Length-ABS(_fPos));
							 END_IF
						END_IF
						stAxis.stPLCTONC.stStartPosition.nRoadID:=stAxis.stNcTOPLC.nCuRoadID;
					ELSE
						IF (_eDirection=E_Direction.DIRECTION_POSITIVE)THEN
							_fDistance:=_fPos-stAxis.stNcTOPLC.fActPos;
						ELSE
							_fDistance:=stAxis.stNcTOPLC.fActPos-_fPos;
						END_IF
					END_IF
				ELSE
					IF(stAxis.stNcTOPLC.nCuRoadID=stAxis.stPLCTONC.nRoadID_2) THEN //第二路段
						
						IF NOT stAxis.stPLCTONC.bRoadDirection  THEN   //正向 
							_fDistance:=_fPos-stAxis.stNcTOPLC.fActPos;
						ELSE
							_fDistance:=stAxis.stNcTOPLC.fActPos-_fPos;
						END_IF
						stAxis.stPLCTONC.stStartPosition.nRoadID:=stAxis.stNcTOPLC.nCuRoadID;
					ELSE
						IF (_eDirection=E_Direction.DIRECTION_POSITIVE)THEN
							_fDistance:=_fPos-stAxis.stNcTOPLC.fActPos;
						ELSE
							_fDistance:=stAxis.stNcTOPLC.fActPos-_fPos;
						END_IF
					END_IF
				END_IF
				
			ELSE
				IF (_eDirection=E_Direction.DIRECTION_POSITIVE)THEN
					_fDistance:=_fPos-stAxis.stNcTOPLC.fActPos;
				ELSE
					_fDistance:=stAxis.stNcTOPLC.fActPos-_fPos;
				END_IF
			END_IF
			_nPathSegment:=1;
	    ELSE
			_nPathSegment:=2;
			_fVeloStart:=stAxis.stNcTOPLC.fActVelo;
			_fVeloEnd:=_fPreTaVel;
			_fTargetVelo:=_fPreTaVel;
			_fDistance:=_fNewAccDis;
			_fAcc:=_fNewAcc;
			_fDec:=_fNewAcc;
			_fPosIn:=_fDealt_S;       
			_fVeloStart_2:=_fPreTaVel;
			_fVeloEnd_2:=0.0;
			_fTargetVelo_2:=_fPreTaVel;
			IF (stAxis.stPLCTONC.nRoadID_2<>0)AND (stAxis.stPLCTONC.nRoadID_1<>0)THEN   //判断指令
				IF (stAxis.stPLCTONC.stStartPosition.nRoadID<>stAxis.stPLCTONC.stEndPosition.nRoadID)THEN
				    IF(stAxis.stNcTOPLC.nCuRoadID=stAxis.stPLCTONC.nRoadID_2) THEN //第二路段
						IF (_eDirection=E_Direction.DIRECTION_POSITIVE)THEN
							 IF NOT stAxis.stPLCTONC.bRoadDirection  THEN   //正向 
								 _fDistance_2:=_fPos-stAxis.stPLCTONC.fRoad1_Length-stAxis.stNcTOPLC.fActPos-_fNewAccDis;
							 ELSE
								 _fDistance_2:=stAxis.stNcTOPLC.fActPos-(stAxis.stPLCTONC.fRoad2_Length-_fPos+stAxis.stPLCTONC.fRoad1_Length)-_fNewAccDis;
							 END_IF
						ELSE
							IF NOT stAxis.stPLCTONC.bRoadDirection  THEN   //正向 
								 _fDistance_2:=ABS(_fPos)-stAxis.stNcTOPLC.fActPos-_fNewAccDis;
							 ELSE
								 _fDistance_2:=stAxis.stNcTOPLC.fActPos-(stAxis.stPLCTONC.fRoad2_Length-ABS(_fPos))-_fNewAccDis;
							 END_IF
						END_IF
						stAxis.stPLCTONC.stStartPosition.nRoadID:=stAxis.stNcTOPLC.nCuRoadID;
					ELSE
						IF (_eDirection=E_Direction.DIRECTION_POSITIVE)THEN
							_fDistance_2:=_fPos-stAxis.stNcTOPLC.fActPos-_fNewAccDis;
						ELSE
							_fDistance_2:=stAxis.stNcTOPLC.fActPos-_fPos-_fNewAccDis;
						END_IF
					END_IF
				ELSE
					IF(stAxis.stNcTOPLC.nCuRoadID=stAxis.stPLCTONC.nRoadID_2) THEN //第二路段
						
						IF NOT stAxis.stPLCTONC.bRoadDirection  THEN   //正向 
							_fDistance_2:=_fPos-stAxis.stNcTOPLC.fActPos-_fNewAccDis;
						ELSE
							_fDistance_2:=stAxis.stNcTOPLC.fActPos-_fPos-_fNewAccDis;
						END_IF
						stAxis.stPLCTONC.stStartPosition.nRoadID:=stAxis.stNcTOPLC.nCuRoadID;
					ELSE
						IF (_eDirection=E_Direction.DIRECTION_POSITIVE)THEN
							_fDistance_2:=_fPos-stAxis.stNcTOPLC.fActPos-_fNewAccDis;
						ELSE
							_fDistance_2:=stAxis.stNcTOPLC.fActPos-_fPos-_fNewAccDis;
						END_IF
					END_IF
				END_IF
				
			ELSE
				IF (_eDirection=E_Direction.DIRECTION_POSITIVE)THEN
					_fDistance_2:=_fPos-stAxis.stNcTOPLC.fActPos-_fNewAccDis;
				ELSE
					_fDistance_2:=stAxis.stNcTOPLC.fActPos-_fPos-_fNewAccDis;
				END_IF
			END_IF
			(*IF (_eDirection=E_Direction.DIRECTION_POSITIVE)THEN
				_fDistance_2:=_fPos-stAxis.stNcTOPLC.fActPos-_fNewAccDis;
			ELSE
				_fDistance_2:=stAxis.stNcTOPLC.fActPos-_fPos-_fNewAccDis;
			END_IF*)
			_fAcc_2:=stAxis.stPLCTONC.stEndPosition.fAccleration;
			_fDec_2:=stAxis.stPLCTONC.stEndPosition.fDeceleration;	
	   END_IF
	
ELSE    
		RETURN;
END_IF
_bSynMode:=TRUE;
_bEnable:=TRUE;
stAxis.stAxisStatus.bSynDecActive:=TRUE;
IF GVL_MC.cDebug  THEN
	_sMessage:=FC_StrContact(stAxis,'next road acc gap control');
	ADSLOGSTR(ADSLOG_MSGTYPE_HINT, _sMessage, '');
END_IF
END_ACTION

ACTION A_NextRoadCatchUp:

//  追击
(***********
   1. 前后动子间距小于防碰撞距离return 
   2. 前后动子间距小于欲减速设置距离，触发减速
   3. 判断当前动子有几段路径，分路径讨论前动子处于路径第几段和处于第几段的加速段、减速段和匀速段

************)
IF (_pNextRoadPremover^.stNcTOPLC.nAxisId<>0)AND (NOT _bSynMode) THEN 
	//预处理减速距离 前瞻距离
	_fDisSet:=0.5*stAxis.stAxisStatus.stPathRef.fTargetVelocity*stAxis.stAxisStatus.stPathRef.fTargetVelocity/_fAcc;        
	
	IF (_nPathSegment=1)THEN 
		IF(_fTime<stAxis.stAxisStatus.stPathRef.aExecutablePath[0].fTa)THEN     // 当前动子处于第一减速段
			
			IF (stAxis.stAxisStatus.stPathRef.aExecutablePath[0].fExpVelo<stAxis.stAxisStatus.stPathRef.aExecutablePath[0].fStartVelo)
				AND (stAxis.stAxisStatus.stPathRef.aExecutablePath[0].fTv<>0)  THEN
				 _fDisSet:=0.5*stAxis.stAxisStatus.stPathRef.aExecutablePath[0].fStartVelo*stAxis.stAxisStatus.stPathRef.aExecutablePath[0].fStartVelo/_fAcc;
			END_IF
			
		END_IF
	ELSIF(_nPathSegment=2)THEN 
		IF(_fTime<stAxis.stAxisStatus.stPathRef.aExecutablePath[0].fTa)THEN
		    _fDisSet:=0.5*stAxis.stAxisStatus.stPathRef.aExecutablePath[0].fStartVelo*stAxis.stAxisStatus.stPathRef.aExecutablePath[0].fStartVelo/_fAcc;
		ELSE
			_fDisSet:=0.5*stAxis.stAxisStatus.stPathRef.aExecutablePath[1].fExpVelo*stAxis.stAxisStatus.stPathRef.aExecutablePath[1].fExpVelo/_fAcc;
		END_IF
	
	ELSE
		;
	END_IF
	_fDealt_S:=_fRealDis-_fGapSet;    //两动子间实时位置偏差，包含gap
	
	IF ((_fRealDis -_fGapSet)<=_fSetDealtGap)AND(_pNextRoadPremover^.stAxisStatus.stPathRef.fTargetVelocity <stAxis.stAxisStatus.stPathRef.fTargetVelocity) THEN    //10.18 
	
		_fPos:=stAxis.stPLCTONC.stEndPosition.fPosition;
		_fTargetVelo:=_pNextRoadPremover^.stAxisStatus.stPathRef.fTargetVelocity;
		_fVeloStart:=stAxis.stNcTOPLC.fActVelo;
		_fVeloEnd:=0;
		_fAcc:=stAxis.stPLCTONC.stEndPosition.fAccleration;
		_fDec:=stAxis.stPLCTONC.stEndPosition.fDeceleration;
		IF (_eDirection=E_Direction.DIRECTION_POSITIVE)THEN
		     _fDistance:=_fPos-stAxis.stNcTOPLC.fActPos;
	    ELSE
			 _fDistance:=stAxis.stNcTOPLC.fActPos-_fPos;
	    END_IF
		_bEnable:=TRUE;
		_nPathSegment:=1;
		stAxis.stAxisStatus.bSynDecActive:=TRUE;
		IF GVL_MC.cDebug  THEN
		     _sMessage:=FC_StrContact(stAxis,'nextroad gap control');
	         ADSLOGSTR(ADSLOG_MSGTYPE_HINT, _sMessage, '');
        END_IF
		
		RETURN;
	 END_IF   //11.22 增加
	
    _fReminDis:=ABS(stAxis.stPLCTONC.stEndPosition.fPosition-stAxis.stNcTOPLC.fActPos);   //剩余目标距离
	
	IF (_fDealt_S-_fDisSet<=0)THEN    //触发减速判断 
		   //IF (_pPremover^.stAxisStatus.stPathRef.fTargetVelocity <stAxis.stAxisStatus.stPathRef.fTargetVelocity) THEN  //11.25注释
		   IF (stAxis.stNcTOPLC.fActVelo>_pNextRoadPremover^.stNcTOPLC.fActVelo) THEN     //11.25修改
			   IF (_fReminDis>_fDisSet)THEN  //判断剩余距离是否满足撞击条件
				    _fPreCurTime:=UDINT_TO_LREAL(_pNextRoadPremover^.stAxisStatus.nNcCycleCounter)*fCycleTime;
			       IF (_pNextRoadPremover^.stAxisStatus.stPathRef._nPathSegmentNum=1)THEN      //判断前动子只有一段路径
					   IF (_fPreCurTime <_pNextRoadPremover^.stAxisStatus.stPathRef.aExecutablePath[0].fTa)THEN      //加速段或减速第一段
						   IF (_pNextRoadPremover^.stAxisStatus.stPathRef.aExecutablePath[0].fExpVelo>_pNextRoadPremover^.stAxisStatus.stPathRef.aExecutablePath[0].fStartVelo)THEN
							   IF (stAxis.stAxisStatus.stPathRef.aExecutablePath[0].fTv<>0) THEN          //加速段
								   A_NextRoadAccSegmengt();
							   END_IF 
						   ELSE    //减速段
							   IF(_pNextRoadPremover^.stAxisStatus.stPathRef.aExecutablePath[0].fTv<>0)THEN 
								   A_NextRoadDecSegment();
							   END_IF
						   END_IF
					   ELSIF (_fPreCurTime <(_pNextRoadPremover^.stAxisStatus.stPathRef.aExecutablePath[0].fTotalTime-_pNextRoadPremover^.stAxisStatus.stPathRef.aExecutablePath[0].fTd))THEN
						   A_NextRoadConVeloSegment();
					   ELSE
						   //
						   RETURN ;  //不处理
					   END_IF
				   //第二段
				   ELSIF(_pNextRoadPremover^.stAxisStatus.stPathRef._nPathSegmentNum=2)THEN
                       IF (_pNextRoadPremover^.stAxisStatus.nSegIndex=0) THEN
						    //IF (_fPreCurTime <_pPremover^.stAxisStatus.stPathRef.aExecutablePath[0].fTa)THEN      //加速段
							IF (_fPreCurTime <_pNextRoadPremover^.stAxisStatus.stPathRef.aExecutablePath[0].fTotalTime)THEN      //减速段  11.29
								A_NextRoadDecSegment_2();
							END_IF
					   ELSIF (_pNextRoadPremover^.stAxisStatus.nSegIndex=1) THEN   //只处理匀速段
						   IF (_fPreCurTime <(_pNextRoadPremover^.stAxisStatus.stPathRef.aExecutablePath[1].fTotalTime-_pNextRoadPremover^.stAxisStatus.stPathRef.aExecutablePath[1].fTd))THEN
						       A_NextRoadConVeloSegment();
						   END_IF   
					   ELSE
						   ;
					   END_IF
					   // 第二段减速段不处理
				   
				   END_IF
			   ELSE
				   RETURN ;
		       END_IF
		   END_IF
	END_IF
END_IF
END_ACTION

ACTION A_NextRoadConVeloSegment:

_fPreTaVel:=_pNextRoadPremover^.stAxisStatus.stPathRef.fTargetVelocity;
_fPreCuVel:=_pNextRoadPremover^.stNcTOPLC.fActVelo;
_fPreAcc:=_fAcc;
_fCuVel:=stAxis.stNcTOPLC.fActVelo;
//_fDealt_S1:=0.5*(_fPreTaVel-_fPreCuVel)*(_fPreTaVel-_fPreCuVel)/_fAcc;
				      
_fNewAcc:=(_fCuVel-_fPreTaVel)*(_fCuVel-_fPreTaVel)*0.5/_fDealt_S;
		   		 
_fDecTime:=	(_fCuVel-_fPreTaVel)/_fNewAcc;
_fNewAccDis:=(_fCuVel*_fCuVel-_fPreTaVel*_fPreTaVel)*0.5/_fNewAcc;
_fMinDis:=_fPreTaVel*_fPreTaVel*0.5/_fPreAcc+_fNewAccDis;

_fPos:=stAxis.stPLCTONC.stEndPosition.fPosition;
	
IF(_fReminDis< _fMinDis)THEN
		_fVeloStart:=stAxis.stNcTOPLC.fActVelo;
	    _fVeloEnd:=0.0;
	    _fTargetVelo:=_pNextRoadPremover^.stAxisStatus.stPathRef.fTargetVelocity;
		IF (stAxis.stPLCTONC.nRoadID_2<>0)AND (stAxis.stPLCTONC.nRoadID_1<>0)THEN   //判断指令
				IF (stAxis.stPLCTONC.stStartPosition.nRoadID<>stAxis.stPLCTONC.stEndPosition.nRoadID)THEN
				    IF(stAxis.stNcTOPLC.nCuRoadID=stAxis.stPLCTONC.nRoadID_2) THEN //第二路段
						IF (_eDirection=E_Direction.DIRECTION_POSITIVE)THEN
							 IF NOT stAxis.stPLCTONC.bRoadDirection  THEN   //正向 
								 _fDistance:=_fPos-stAxis.stPLCTONC.fRoad1_Length-stAxis.stNcTOPLC.fActPos;
							 ELSE
								 _fDistance:=stAxis.stNcTOPLC.fActPos-(stAxis.stPLCTONC.fRoad2_Length-_fPos+stAxis.stPLCTONC.fRoad1_Length);
							 END_IF
						ELSE
							IF NOT stAxis.stPLCTONC.bRoadDirection  THEN   //正向 
								 _fDistance:=ABS(_fPos)-stAxis.stNcTOPLC.fActPos;
							 ELSE
								 _fDistance:=stAxis.stNcTOPLC.fActPos-(stAxis.stPLCTONC.fRoad2_Length-ABS(_fPos));
							 END_IF
						END_IF
						stAxis.stPLCTONC.stStartPosition.nRoadID:=stAxis.stNcTOPLC.nCuRoadID;
					ELSE
						IF (_eDirection=E_Direction.DIRECTION_POSITIVE)THEN
							_fDistance:=_fPos-stAxis.stNcTOPLC.fActPos;
						ELSE
							_fDistance:=stAxis.stNcTOPLC.fActPos-_fPos;
						END_IF
					END_IF
				ELSE
					IF(stAxis.stNcTOPLC.nCuRoadID=stAxis.stPLCTONC.nRoadID_2) THEN //第二路段
						
						IF NOT stAxis.stPLCTONC.bRoadDirection  THEN   //正向 
							_fDistance:=_fPos-stAxis.stNcTOPLC.fActPos;
						ELSE
							_fDistance:=stAxis.stNcTOPLC.fActPos-_fPos;
						END_IF
						stAxis.stPLCTONC.stStartPosition.nRoadID:=stAxis.stNcTOPLC.nCuRoadID;
					ELSE
						IF (_eDirection=E_Direction.DIRECTION_POSITIVE)THEN
							_fDistance:=_fPos-stAxis.stNcTOPLC.fActPos;
						ELSE
							_fDistance:=stAxis.stNcTOPLC.fActPos-_fPos;
						END_IF
					END_IF
				END_IF
				
		ELSE
				IF (_eDirection=E_Direction.DIRECTION_POSITIVE)THEN
					_fDistance:=_fPos-stAxis.stNcTOPLC.fActPos;
				ELSE
					_fDistance:=stAxis.stNcTOPLC.fActPos-_fPos;
				END_IF
		END_IF
		(*IF (_eDirection=E_Direction.DIRECTION_POSITIVE)THEN
			_fDistance:=_fPos-stAxis.stNcTOPLC.fActPos;
		ELSE
			_fDistance:=stAxis.stNcTOPLC.fActPos-_fPos;
		END_IF*)
		_fAcc:=stAxis.stPLCTONC.stEndPosition.fAccleration;
	    _fDec:=stAxis.stPLCTONC.stEndPosition.fDeceleration;
		_nPathSegment:=1;
ELSE
		_nPathSegment:=2;
		_fVeloStart:=stAxis.stNcTOPLC.fActVelo;
	    _fVeloEnd:=_fPreTaVel;
	    _fTargetVelo:=_fPreTaVel;
		_fDistance:=_fNewAccDis;
		_fAcc:=_fNewAcc;
	    _fDec:=_fNewAcc;
		_fPosIn:=_fDealt_S;       //11.29
	    _fVeloStart_2:=_fPreTaVel;
	    _fVeloEnd_2:=0.0;
	    _fTargetVelo_2:=_fPreTaVel;
		IF (stAxis.stPLCTONC.nRoadID_2<>0)AND (stAxis.stPLCTONC.nRoadID_1<>0)THEN   //判断指令
				IF (stAxis.stPLCTONC.stStartPosition.nRoadID<>stAxis.stPLCTONC.stEndPosition.nRoadID)THEN
				    IF(stAxis.stNcTOPLC.nCuRoadID=stAxis.stPLCTONC.nRoadID_2) THEN //第二路段
						IF (_eDirection=E_Direction.DIRECTION_POSITIVE)THEN
							 IF NOT stAxis.stPLCTONC.bRoadDirection  THEN   //正向 
								 _fDistance_2:=_fPos-stAxis.stPLCTONC.fRoad1_Length-stAxis.stNcTOPLC.fActPos-_fNewAccDis;
							 ELSE
								 _fDistance_2:=stAxis.stNcTOPLC.fActPos-(stAxis.stPLCTONC.fRoad2_Length-_fPos+stAxis.stPLCTONC.fRoad1_Length)-_fNewAccDis;
							 END_IF
						ELSE
							IF NOT stAxis.stPLCTONC.bRoadDirection  THEN   //正向 
								 _fDistance_2:=ABS(_fPos)-stAxis.stNcTOPLC.fActPos-_fNewAccDis;
							 ELSE
								 _fDistance_2:=stAxis.stNcTOPLC.fActPos-(stAxis.stPLCTONC.fRoad2_Length-ABS(_fPos))-_fNewAccDis;
							 END_IF
						END_IF
						stAxis.stPLCTONC.stStartPosition.nRoadID:=stAxis.stNcTOPLC.nCuRoadID;
					ELSE
						IF (_eDirection=E_Direction.DIRECTION_POSITIVE)THEN
							_fDistance_2:=_fPos-stAxis.stNcTOPLC.fActPos-_fNewAccDis;
						ELSE
							_fDistance_2:=stAxis.stNcTOPLC.fActPos-_fPos-_fNewAccDis;
						END_IF
					END_IF
				ELSE
					IF(stAxis.stNcTOPLC.nCuRoadID=stAxis.stPLCTONC.nRoadID_2) THEN //第二路段
						
						IF NOT stAxis.stPLCTONC.bRoadDirection  THEN   //正向 
							_fDistance_2:=_fPos-stAxis.stNcTOPLC.fActPos-_fNewAccDis;
						ELSE
							_fDistance_2:=stAxis.stNcTOPLC.fActPos-_fPos-_fNewAccDis;
						END_IF
						stAxis.stPLCTONC.stStartPosition.nRoadID:=stAxis.stNcTOPLC.nCuRoadID;
					ELSE
						IF (_eDirection=E_Direction.DIRECTION_POSITIVE)THEN
							_fDistance_2:=_fPos-stAxis.stNcTOPLC.fActPos-_fNewAccDis;
						ELSE
							_fDistance_2:=stAxis.stNcTOPLC.fActPos-_fPos-_fNewAccDis;
						END_IF
					END_IF
				END_IF
				
			ELSE
				IF (_eDirection=E_Direction.DIRECTION_POSITIVE)THEN
					_fDistance_2:=_fPos-stAxis.stNcTOPLC.fActPos-_fNewAccDis;
				ELSE
					_fDistance_2:=stAxis.stNcTOPLC.fActPos-_fPos-_fNewAccDis;
				END_IF
			END_IF
		(*IF (_eDirection=E_Direction.DIRECTION_POSITIVE)THEN
			_fDistance_2:=_fPos-stAxis.stNcTOPLC.fActPos-_fNewAccDis;
		ELSE
			_fDistance_2:=stAxis.stNcTOPLC.fActPos-_fPos-_fNewAccDis;
		END_IF*)
		_fAcc_2:=stAxis.stPLCTONC.stEndPosition.fAccleration;
	    _fDec_2:=stAxis.stPLCTONC.stEndPosition.fDeceleration;
END_IF

_bSynMode:=TRUE;
_bEnable:=TRUE;
stAxis.stAxisStatus.bSynDecActive:=TRUE;
IF GVL_MC.cDebug  THEN
		     _sMessage:=FC_StrContact(stAxis,'next road con gap control');
	         ADSLOGSTR(ADSLOG_MSGTYPE_HINT, _sMessage, '');
END_IF
END_ACTION

ACTION A_NextRoadDecSegment:

_fPreTaVel:=_pNextRoadPremover^.stAxisStatus.stPathRef.fTargetVelocity;
_fPreCuVel:=_pNextRoadPremover^.stNcTOPLC.fActVelo;
_fPreAcc:=_fAcc;
_fCuVel:=stAxis.stNcTOPLC.fActVelo;
// 计算前动子的减速距离
_fPre_S:=(_fPreCuVel-_fPreTaVel)*(_fPreCuVel-_fPreTaVel)*0.5/_pNextRoadPremover^.stAxisStatus.stPathRef.aExecutablePath[0].fDeceleration;
		      	   
//_fNewAcc:=(_fCuVel-_fPreTaVel)*(_fCuVel-_fPreTaVel)*0.5/_fDealt_S;  //06.18 
_fNewAcc:=(_fCuVel-_fPreTaVel)*(_fCuVel-_fPreTaVel)*0.5/(_fDealt_S+_fPre_S);  //06.18		      	   
//_fNewAcc:=(_fCuVel-_fPreTaVel)*(_fCuVel-_fPreTaVel)*0.5/_fDealt_S;
_fDecTime:=	(_fCuVel-_fPreTaVel)/_fNewAcc;
_fNewAccDis:=(_fCuVel*_fCuVel-_fPreTaVel*_fPreTaVel)*0.5/_fNewAcc;
_fMinDis:=_fPreTaVel*_fPreTaVel*0.5/_fPreAcc+_fNewAccDis;

_fPos:=stAxis.stPLCTONC.stEndPosition.fPosition;

IF(_fReminDis< _fMinDis)THEN
		_fVeloStart:=stAxis.stNcTOPLC.fActVelo;
	    _fVeloEnd:=0.0;
	    _fTargetVelo:=_pNextRoadPremover^.stAxisStatus.stPathRef.fTargetVelocity;
		IF (stAxis.stPLCTONC.nRoadID_2<>0)AND (stAxis.stPLCTONC.nRoadID_1<>0)THEN   //判断指令
				IF (stAxis.stPLCTONC.stStartPosition.nRoadID<>stAxis.stPLCTONC.stEndPosition.nRoadID)THEN
				    IF(stAxis.stNcTOPLC.nCuRoadID=stAxis.stPLCTONC.nRoadID_2) THEN //第二路段
						IF (_eDirection=E_Direction.DIRECTION_POSITIVE)THEN
							 IF NOT stAxis.stPLCTONC.bRoadDirection  THEN   //正向 
								 _fDistance:=_fPos-stAxis.stPLCTONC.fRoad1_Length-stAxis.stNcTOPLC.fActPos;
							 ELSE
								 _fDistance:=stAxis.stNcTOPLC.fActPos-(stAxis.stPLCTONC.fRoad2_Length-_fPos+stAxis.stPLCTONC.fRoad1_Length);
							 END_IF
						ELSE
							IF NOT stAxis.stPLCTONC.bRoadDirection  THEN   //正向 
								 _fDistance:=ABS(_fPos)-stAxis.stNcTOPLC.fActPos;
							 ELSE
								 _fDistance:=stAxis.stNcTOPLC.fActPos-(stAxis.stPLCTONC.fRoad2_Length-ABS(_fPos));
							 END_IF
						END_IF
						stAxis.stPLCTONC.stStartPosition.nRoadID:=stAxis.stNcTOPLC.nCuRoadID;
					ELSE
						IF (_eDirection=E_Direction.DIRECTION_POSITIVE)THEN
							_fDistance:=_fPos-stAxis.stNcTOPLC.fActPos;
						ELSE
							_fDistance:=stAxis.stNcTOPLC.fActPos-_fPos;
						END_IF
					END_IF
				ELSE
					IF(stAxis.stNcTOPLC.nCuRoadID=stAxis.stPLCTONC.nRoadID_2) THEN //第二路段
						
						IF NOT stAxis.stPLCTONC.bRoadDirection  THEN   //正向 
							_fDistance:=_fPos-stAxis.stNcTOPLC.fActPos;
						ELSE
							_fDistance:=stAxis.stNcTOPLC.fActPos-_fPos;
						END_IF
						stAxis.stPLCTONC.stStartPosition.nRoadID:=stAxis.stNcTOPLC.nCuRoadID;
					ELSE
						IF (_eDirection=E_Direction.DIRECTION_POSITIVE)THEN
							_fDistance:=_fPos-stAxis.stNcTOPLC.fActPos;
						ELSE
							_fDistance:=stAxis.stNcTOPLC.fActPos-_fPos;
						END_IF
					END_IF
				END_IF
				
		ELSE
				IF (_eDirection=E_Direction.DIRECTION_POSITIVE)THEN
					_fDistance:=_fPos-stAxis.stNcTOPLC.fActPos;
				ELSE
					_fDistance:=stAxis.stNcTOPLC.fActPos-_fPos;
				END_IF
		END_IF
		(*IF (_eDirection=E_Direction.DIRECTION_POSITIVE)THEN
			_fDistance:=_fPos-stAxis.stNcTOPLC.fActPos;
		ELSE
			_fDistance:=stAxis.stNcTOPLC.fActPos-_fPos;
		END_IF*)
		_fAcc:=stAxis.stPLCTONC.stEndPosition.fAccleration;
	    _fDec:=stAxis.stPLCTONC.stEndPosition.fDeceleration;
		_nPathSegment:=1;
ELSE
		_nPathSegment:=2;
		_fVeloStart:=stAxis.stNcTOPLC.fActVelo;
	    _fVeloEnd:=_fPreTaVel;
	    _fTargetVelo:=_fPreTaVel;
		_fDistance:=_fNewAccDis;
		_fAcc:=_fNewAcc;
	    _fDec:=_fNewAcc;
		
	    _fVeloStart_2:=_fPreTaVel;
	    _fVeloEnd_2:=0.0;
	    _fTargetVelo_2:=_fPreTaVel;
		_fPosIn:=_fDealt_S;       // 25.01.17
		IF (stAxis.stPLCTONC.nRoadID_2<>0)AND (stAxis.stPLCTONC.nRoadID_1<>0)THEN   //判断指令
				IF (stAxis.stPLCTONC.stStartPosition.nRoadID<>stAxis.stPLCTONC.stEndPosition.nRoadID)THEN
				    IF(stAxis.stNcTOPLC.nCuRoadID=stAxis.stPLCTONC.nRoadID_2) THEN //第二路段
						IF (_eDirection=E_Direction.DIRECTION_POSITIVE)THEN
							 IF NOT stAxis.stPLCTONC.bRoadDirection  THEN   //正向 
								 _fDistance_2:=_fPos-stAxis.stPLCTONC.fRoad1_Length-stAxis.stNcTOPLC.fActPos-_fNewAccDis;
							 ELSE
								 _fDistance_2:=stAxis.stNcTOPLC.fActPos-(stAxis.stPLCTONC.fRoad2_Length-_fPos+stAxis.stPLCTONC.fRoad1_Length)-_fNewAccDis;
							 END_IF
						ELSE
							IF NOT stAxis.stPLCTONC.bRoadDirection  THEN   //正向 
								 _fDistance_2:=ABS(_fPos)-stAxis.stNcTOPLC.fActPos-_fNewAccDis;
							 ELSE
								 _fDistance_2:=stAxis.stNcTOPLC.fActPos-(stAxis.stPLCTONC.fRoad2_Length-ABS(_fPos))-_fNewAccDis;
							 END_IF
						END_IF
						stAxis.stPLCTONC.stStartPosition.nRoadID:=stAxis.stNcTOPLC.nCuRoadID;
					ELSE
						IF (_eDirection=E_Direction.DIRECTION_POSITIVE)THEN
							_fDistance_2:=_fPos-stAxis.stNcTOPLC.fActPos-_fNewAccDis;
						ELSE
							_fDistance_2:=stAxis.stNcTOPLC.fActPos-_fPos-_fNewAccDis;
						END_IF
					END_IF
				ELSE
					IF(stAxis.stNcTOPLC.nCuRoadID=stAxis.stPLCTONC.nRoadID_2) THEN //第二路段
						
						IF NOT stAxis.stPLCTONC.bRoadDirection  THEN   //正向 
							_fDistance_2:=_fPos-stAxis.stNcTOPLC.fActPos-_fNewAccDis;
						ELSE
							_fDistance_2:=stAxis.stNcTOPLC.fActPos-_fPos-_fNewAccDis;
						END_IF
						stAxis.stPLCTONC.stStartPosition.nRoadID:=stAxis.stNcTOPLC.nCuRoadID;
					ELSE
						IF (_eDirection=E_Direction.DIRECTION_POSITIVE)THEN
							_fDistance_2:=_fPos-stAxis.stNcTOPLC.fActPos-_fNewAccDis;
						ELSE
							_fDistance_2:=stAxis.stNcTOPLC.fActPos-_fPos-_fNewAccDis;
						END_IF
					END_IF
				END_IF
				
		ELSE
				IF (_eDirection=E_Direction.DIRECTION_POSITIVE)THEN
					_fDistance_2:=_fPos-stAxis.stNcTOPLC.fActPos-_fNewAccDis;
				ELSE
					_fDistance_2:=stAxis.stNcTOPLC.fActPos-_fPos-_fNewAccDis;
				END_IF
		END_IF
		(*IF (_eDirection=E_Direction.DIRECTION_POSITIVE)THEN
			_fDistance_2:=_fPos-stAxis.stNcTOPLC.fActPos-_fNewAccDis;
		ELSE
			_fDistance_2:=stAxis.stNcTOPLC.fActPos-_fPos-_fNewAccDis;
		END_IF*)
		_fAcc_2:=stAxis.stPLCTONC.stEndPosition.fAccleration;
	    _fDec_2:=stAxis.stPLCTONC.stEndPosition.fDeceleration;
END_IF
_bSynMode:=TRUE;
_bEnable:=TRUE;
stAxis.stAxisStatus.bSynDecActive:=TRUE;

IF GVL_MC.cDebug  THEN
		     _sMessage:=FC_StrContact(stAxis,'next road dec gap control');
	         ADSLOGSTR(ADSLOG_MSGTYPE_HINT, _sMessage, '');
END_IF
END_ACTION

ACTION A_NextRoadDecSegment_2:

_fPreTaVel:=_pNextRoadPremover^.stAxisStatus.stPathRef.fTargetVelocity;
_fPreCuVel:=_pNextRoadPremover^.stNcTOPLC.fActVelo;
_fPreAcc:=_fAcc;
_fCuVel:=stAxis.stNcTOPLC.fActVelo;

//_fPreDealt_S:=0.5*(_pPremover^.stAxisStatus.stPathRef.aExecutablePath[0].fTa-_fPreCurTime)*_fPreCuVel;
//_fPreDealt_S:=_pPremover^.stAxisStatus.stPathRef.fDealtInPos- 0.5*(_fPreTaVel+_fPreCuVel)*_fPreCurTime; //11.29	

 _fPreSeg1TotalTime :=_pNextRoadPremover^.stAxisStatus.stPathRef.aExecutablePath[0].fTotalTime;   //05.26
//_fPreDealt_S:=0.5*(_pPremover^.stAxisStatus.stPathRef.aExecutablePath[0].fTa-_fPreCurTime)*_fPreCuVel;
//_fPreDealt_S:=_pPremover^.stAxisStatus.stPathRef.fDealtInPos- 0.5*(_fPreTaVel+_fPreCuVel)*_fPreCurTime; //05.26  
_fPreDealt_S:=0.5*(_fPreCuVel-_fPreTaVel)*( _fPreSeg1TotalTime-_fPreCurTime); //05.26 			      	   
_fNewAcc:=(_fCuVel-_fPreTaVel)*(_fCuVel-_fPreTaVel)*0.5/(_fDealt_S+_fPreDealt_S);
		   		 
_fDecTime:=	(_fCuVel-_fPreTaVel)/_fNewAcc;
_fNewAccDis:=(_fCuVel*_fCuVel-_fPreTaVel*_fPreTaVel)*0.5/_fNewAcc;

_fMinDis:=_fPreTaVel*_fPreTaVel*0.5/_fPreAcc+_fNewAccDis;

_fPos:=stAxis.stPLCTONC.stEndPosition.fPosition;

IF( _fReminDis< _fMinDis)THEN
		_fVeloStart:=stAxis.stNcTOPLC.fActVelo;
	    _fVeloEnd:=0.0;
	    _fTargetVelo:=_pNextRoadPremover^.stAxisStatus.stPathRef.fTargetVelocity;
		IF (stAxis.stPLCTONC.nRoadID_2<>0)AND (stAxis.stPLCTONC.nRoadID_1<>0)THEN   //判断指令
				IF (stAxis.stPLCTONC.stStartPosition.nRoadID<>stAxis.stPLCTONC.stEndPosition.nRoadID)THEN
				    IF(stAxis.stNcTOPLC.nCuRoadID=stAxis.stPLCTONC.nRoadID_2) THEN //第二路段
						IF (_eDirection=E_Direction.DIRECTION_POSITIVE)THEN
							 IF NOT stAxis.stPLCTONC.bRoadDirection  THEN   //正向 
								 _fDistance:=_fPos-stAxis.stPLCTONC.fRoad1_Length-stAxis.stNcTOPLC.fActPos;
							 ELSE
								 _fDistance:=stAxis.stNcTOPLC.fActPos-(stAxis.stPLCTONC.fRoad2_Length-_fPos+stAxis.stPLCTONC.fRoad1_Length);
							 END_IF
						ELSE
							IF NOT stAxis.stPLCTONC.bRoadDirection  THEN   //正向 
								 _fDistance:=ABS(_fPos)-stAxis.stNcTOPLC.fActPos;
							 ELSE
								 _fDistance:=stAxis.stNcTOPLC.fActPos-(stAxis.stPLCTONC.fRoad2_Length-ABS(_fPos));
							 END_IF
						END_IF
						stAxis.stPLCTONC.stStartPosition.nRoadID:=stAxis.stNcTOPLC.nCuRoadID;
					ELSE
						IF (_eDirection=E_Direction.DIRECTION_POSITIVE)THEN
							_fDistance:=_fPos-stAxis.stNcTOPLC.fActPos;
						ELSE
							_fDistance:=stAxis.stNcTOPLC.fActPos-_fPos;
						END_IF
					END_IF
				ELSE
					IF(stAxis.stNcTOPLC.nCuRoadID=stAxis.stPLCTONC.nRoadID_2) THEN //第二路段
						
						IF NOT stAxis.stPLCTONC.bRoadDirection  THEN   //正向 
							_fDistance:=_fPos-stAxis.stNcTOPLC.fActPos;
						ELSE
							_fDistance:=stAxis.stNcTOPLC.fActPos-_fPos;
						END_IF
						stAxis.stPLCTONC.stStartPosition.nRoadID:=stAxis.stNcTOPLC.nCuRoadID;
					ELSE
						IF (_eDirection=E_Direction.DIRECTION_POSITIVE)THEN
							_fDistance:=_fPos-stAxis.stNcTOPLC.fActPos;
						ELSE
							_fDistance:=stAxis.stNcTOPLC.fActPos-_fPos;
						END_IF
					END_IF
				END_IF
				
